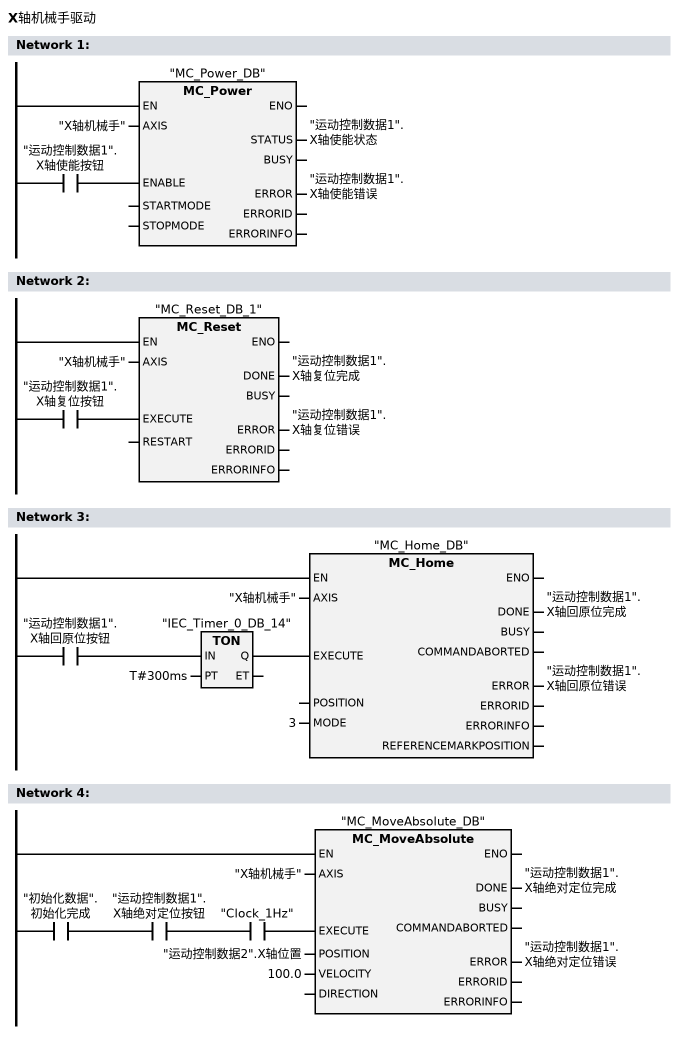
   "MC_Power_DB"(Axis := "X轴机械手",   // MC_Power
                 Enable := "运动控制数据1".X轴使能按钮,
                 Status => "运动控制数据1".X轴使能状态,
                 Error => "运动控制数据1".X轴使能错误);
END_REGION

REGION Network 2
   "MC_Reset_DB_1"(Axis := "X轴机械手",   // MC_Reset
                   Execute := "运动控制数据1".X轴复位按钮,
                   Done => "运动控制数据1".X轴复位完成,
                   Error => "运动控制数据1".X轴复位错误);
END_REGION

REGION Network 3
   "IEC_Timer_0_DB_14".TON(IN := "运动控制数据1".X轴回原位按钮, PT := T#300ms);
   "MC_Home_DB"(Axis := "X轴机械手",   // MC_Home
                Execute := "IEC_Timer_0_DB_14".Q,
                Mode := 3,
                Done => "运动控制数据1".X轴回原位完成,
                Error => "运动控制数据1".X轴回原位错误);
END_REGION

REGION Network 4
   "MC_MoveAbsolute_DB"(Axis := "X轴机械手",   // MC_MoveAbsolute
                        Execute := "初始化数据".初始化完成 AND "运动控制数据1".X轴绝对定位按钮 AND "Clock_1Hz",
                        Position := "运动控制数据2".X轴位置,
                        Velocity := 100.0,
                        Done => "运动控制数据1".X轴绝对定位完成,
                        Error => "运动控制数据1".X轴绝对定位错误);
END_REGION
END_FUNCTION

FUNCTION "Y轴机械手驱动" : Void   // FC2, LAD
{ S7_Optimized_Access := 'TRUE' }
VERSION : 0.1
BEGIN

REGION Network 1
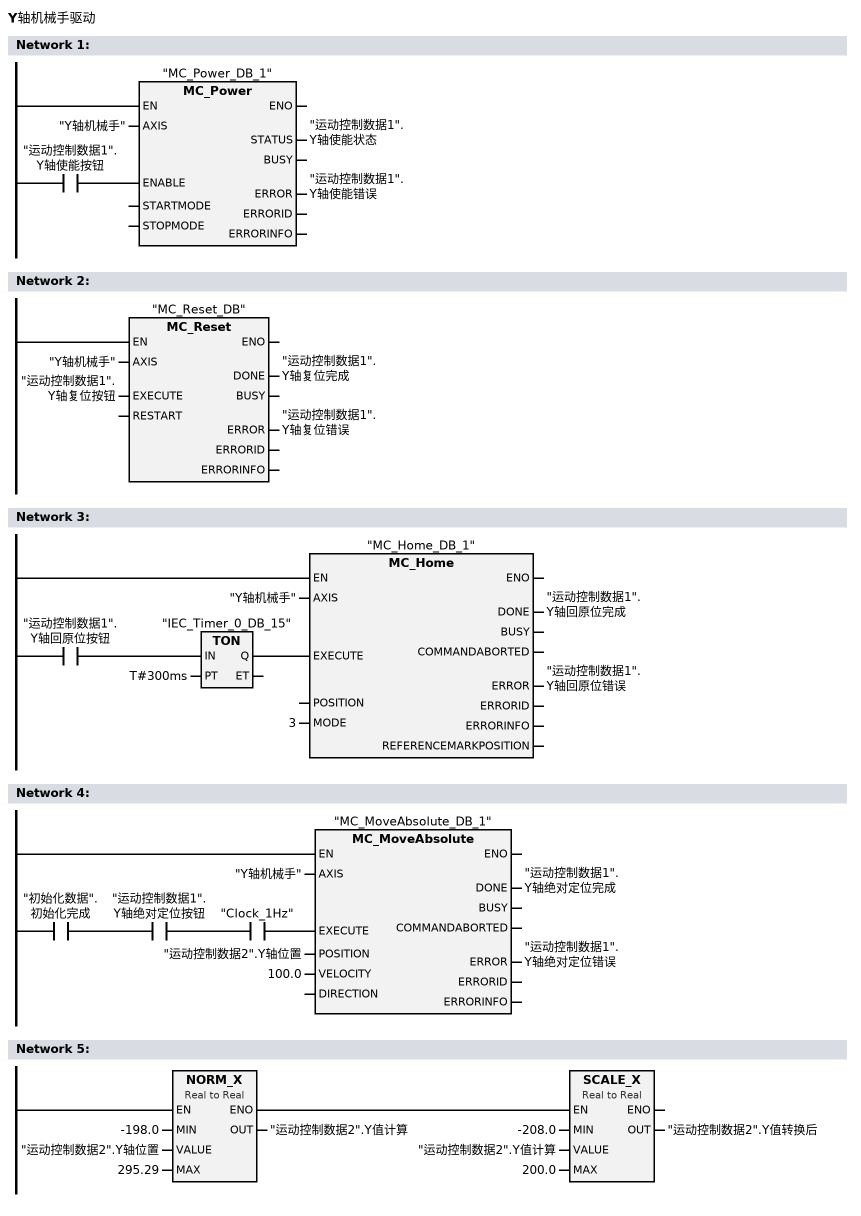
   "MC_Power_DB_1"(Axis := "Y轴机械手",   // MC_Power
                   Enable := "运动控制数据1".Y轴使能按钮,
                   Status => "运动控制数据1".Y轴使能状态,
                   Error => "运动控制数据1".Y轴使能错误);
END_REGION

REGION Network 2
   "MC_Reset_DB"(Axis := "Y轴机械手",   // MC_Reset
                 Execute := "运动控制数据1".Y轴复位按钮,
                 Done => "运动控制数据1".Y轴复位完成,
                 Error => "运动控制数据1".Y轴复位错误);
END_REGION

REGION Network 3
   "IEC_Timer_0_DB_15".TON(IN := "运动控制数据1".Y轴回原位按钮, PT := T#300ms);
   "MC_Home_DB_1"(Axis := "Y轴机械手",   // MC_Home
                  Execute := "IEC_Timer_0_DB_15".Q,
                  Mode := 3,
                  Done => "运动控制数据1".Y轴回原位完成,
                  Error => "运动控制数据1".Y轴回原位错误);
END_REGION

REGION Network 4
   "MC_MoveAbsolute_DB_1"(Axis := "Y轴机械手",   // MC_MoveAbsolute
                          Execute := "初始化数据".初始化完成 AND "运动控制数据1".Y轴绝对定位按钮 AND "Clock_1Hz",
                          Position := "运动控制数据2".Y轴位置,
                          Velocity := 100.0,
                          Done => "运动控制数据1".Y轴绝对定位完成,
                          Error => "运动控制数据1".Y轴绝对定位错误);
END_REGION

REGION Network 5
   RUNG wire#powerrail
      { S7_Templates := "[SrcType := Real, DestType := Real]" } Normalize(min := -198.0, value := "运动控制数据2".Y轴位置, max := 295.29, out => "运动控制数据2".Y值计算)
      { S7_Templates := "[SrcType := Real, DestType := Real]" } Scale(min := -208.0, value := "运动控制数据2".Y值计算, max := 200.0, out => "运动控制数据2".Y值转换后)
   END_RUNG
   // the same network as SCL:
   "运动控制数据2".Y值计算 := NORM_X(MIN := -198.0, VALUE := "运动控制数据2".Y轴位置, MAX := 295.29);
   "运动控制数据2".Y值转换后 := SCALE_X(MIN := -208.0, VALUE := "运动控制数据2".Y值计算, MAX := 200.0);
END_REGION
END_FUNCTION

FUNCTION "传输皮带" : Void   // FC3, LAD
{ S7_Optimized_Access := 'TRUE' }
VERSION : 0.1
BEGIN

REGION Network 1
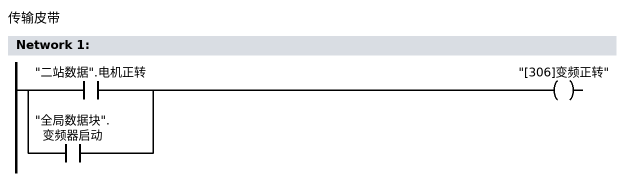
   RUNG wire#powerrail
      Contact( "二站数据".电机正转 )
      wire#w1
      Coil( "[306]变频正转" )
   END_RUNG
   RUNG wire#powerrail
      Contact( "全局数据块".变频器启动 )
   END_RUNG wire#w1
   // the same network as SCL:
   "[306]变频正转" := "二站数据".电机正转 OR "全局数据块".变频器启动;
END_REGION
END_FUNCTION

FUNCTION "00.轴初始化程序" : Void   // FC11, LAD
{ S7_Optimized_Access := 'TRUE' }
VERSION : 0.1
   VAR_TEMP   // added for the SCL form of the ladder/FBD networks
      _w1 : Bool;
   END_VAR
BEGIN

REGION Network 1
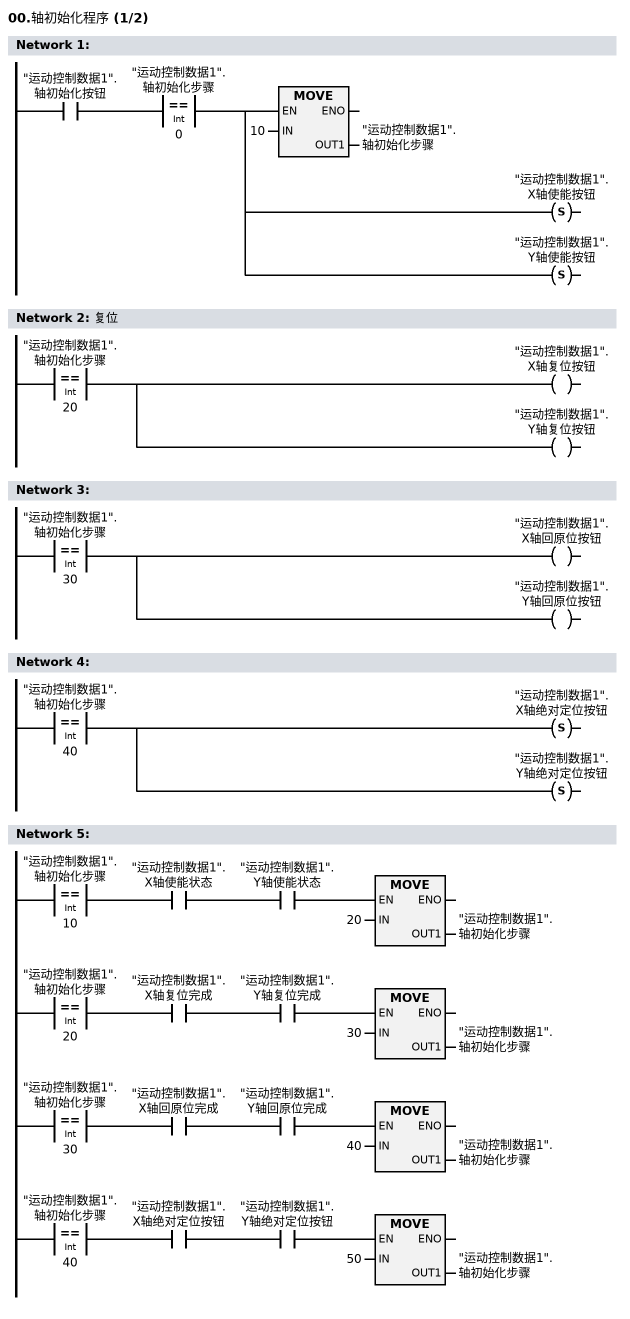
   RUNG wire#powerrail
      Contact( "运动控制数据1".轴初始化按钮 )
      { S7_Templates := "SrcType := Int" } EQ_Contact(in1 := "运动控制数据1".轴初始化步骤, in2 := 0)
      wire#w1
      Move(in := 10, out1 => "运动控制数据1".轴初始化步骤)
   END_RUNG
   RUNG wire#w1
      S_Coil( "运动控制数据1".X轴使能按钮 )
   END_RUNG
   RUNG wire#w1
      S_Coil( "运动控制数据1".Y轴使能按钮 )
   END_RUNG
   // the same network as SCL:
   #_w1 := "运动控制数据1".轴初始化按钮 AND ("运动控制数据1".轴初始化步骤 = 0);
   IF #_w1 THEN
       "运动控制数据1".轴初始化步骤 := 10;
       "运动控制数据1".X轴使能按钮 := TRUE;
       "运动控制数据1".Y轴使能按钮 := TRUE;
   END_IF;
END_REGION

REGION Network 2: 复位
   RUNG wire#powerrail
      { S7_Templates := "SrcType := Int" } EQ_Contact(in1 := "运动控制数据1".轴初始化步骤, in2 := 20)
      wire#w1
      Coil( "运动控制数据1".X轴复位按钮 )
   END_RUNG
   RUNG wire#w1
      Coil( "运动控制数据1".Y轴复位按钮 )
   END_RUNG
   // the same network as SCL:
   "运动控制数据1".X轴复位按钮 := "运动控制数据1".轴初始化步骤 = 20;
   "运动控制数据1".Y轴复位按钮 := "运动控制数据1".X轴复位按钮;
END_REGION

REGION Network 3
   RUNG wire#powerrail
      { S7_Templates := "SrcType := Int" } EQ_Contact(in1 := "运动控制数据1".轴初始化步骤, in2 := 30)
      wire#w1
      Coil( "运动控制数据1".X轴回原位按钮 )
   END_RUNG
   RUNG wire#w1
      Coil( "运动控制数据1".Y轴回原位按钮 )
   END_RUNG
   // the same network as SCL:
   "运动控制数据1".X轴回原位按钮 := "运动控制数据1".轴初始化步骤 = 30;
   "运动控制数据1".Y轴回原位按钮 := "运动控制数据1".X轴回原位按钮;
END_REGION

REGION Network 4
   RUNG wire#powerrail
      { S7_Templates := "SrcType := Int" } EQ_Contact(in1 := "运动控制数据1".轴初始化步骤, in2 := 40)
      wire#w1
      S_Coil( "运动控制数据1".X轴绝对定位按钮 )
   END_RUNG
   RUNG wire#w1
      S_Coil( "运动控制数据1".Y轴绝对定位按钮 )
   END_RUNG
   // the same network as SCL:
   IF "运动控制数据1".轴初始化步骤 = 40 THEN
       "运动控制数据1".X轴绝对定位按钮 := TRUE;
       "运动控制数据1".Y轴绝对定位按钮 := TRUE;
   END_IF;
END_REGION

REGION Network 5
   RUNG wire#powerrail
      { S7_Templates := "SrcType := Int" } EQ_Contact(in1 := "运动控制数据1".轴初始化步骤, in2 := 10)
      Contact( "运动控制数据1".X轴使能状态 )
      Contact( "运动控制数据1".Y轴使能状态 )
      Move(in := 20, out1 => "运动控制数据1".轴初始化步骤)
   END_RUNG
   RUNG wire#powerrail
      { S7_Templates := "SrcType := Int" } EQ_Contact(in1 := "运动控制数据1".轴初始化步骤, in2 := 20)
      Contact( "运动控制数据1".X轴复位完成 )
      Contact( "运动控制数据1".Y轴复位完成 )
      Move(in := 30, out1 => "运动控制数据1".轴初始化步骤)
   END_RUNG
   RUNG wire#powerrail
      { S7_Templates := "SrcType := Int" } EQ_Contact(in1 := "运动控制数据1".轴初始化步骤, in2 := 30)
      Contact( "运动控制数据1".X轴回原位完成 )
      Contact( "运动控制数据1".Y轴回原位完成 )
      Move(in := 40, out1 => "运动控制数据1".轴初始化步骤)
   END_RUNG
   RUNG wire#powerrail
      { S7_Templates := "SrcType := Int" } EQ_Contact(in1 := "运动控制数据1".轴初始化步骤, in2 := 40)
      Contact( "运动控制数据1".X轴绝对定位按钮 )
      Contact( "运动控制数据1".Y轴绝对定位按钮 )
      Move(in := 50, out1 => "运动控制数据1".轴初始化步骤)
   END_RUNG
   // the same network as SCL:
   IF ("运动控制数据1".轴初始化步骤 = 10) AND "运动控制数据1".X轴使能状态 AND "运动控制数据1".Y轴使能状态 THEN "运动控制数据1".轴初始化步骤 := 20; END_IF;
   IF ("运动控制数据1".轴初始化步骤 = 20) AND "运动控制数据1".X轴复位完成 AND "运动控制数据1".Y轴复位完成 THEN "运动控制数据1".轴初始化步骤 := 30; END_IF;
   IF ("运动控制数据1".轴初始化步骤 = 30) AND "运动控制数据1".X轴回原位完成 AND "运动控制数据1".Y轴回原位完成 THEN
       "运动控制数据1".轴初始化步骤 := 40;
   END_IF;
   IF ("运动控制数据1".轴初始化步骤 = 40) AND "运动控制数据1".X轴绝对定位按钮 AND "运动控制数据1".Y轴绝对定位按钮 THEN
       "运动控制数据1".轴初始化步骤 := 50;
   END_IF;
END_REGION

REGION Network 6: 轴初始化完成
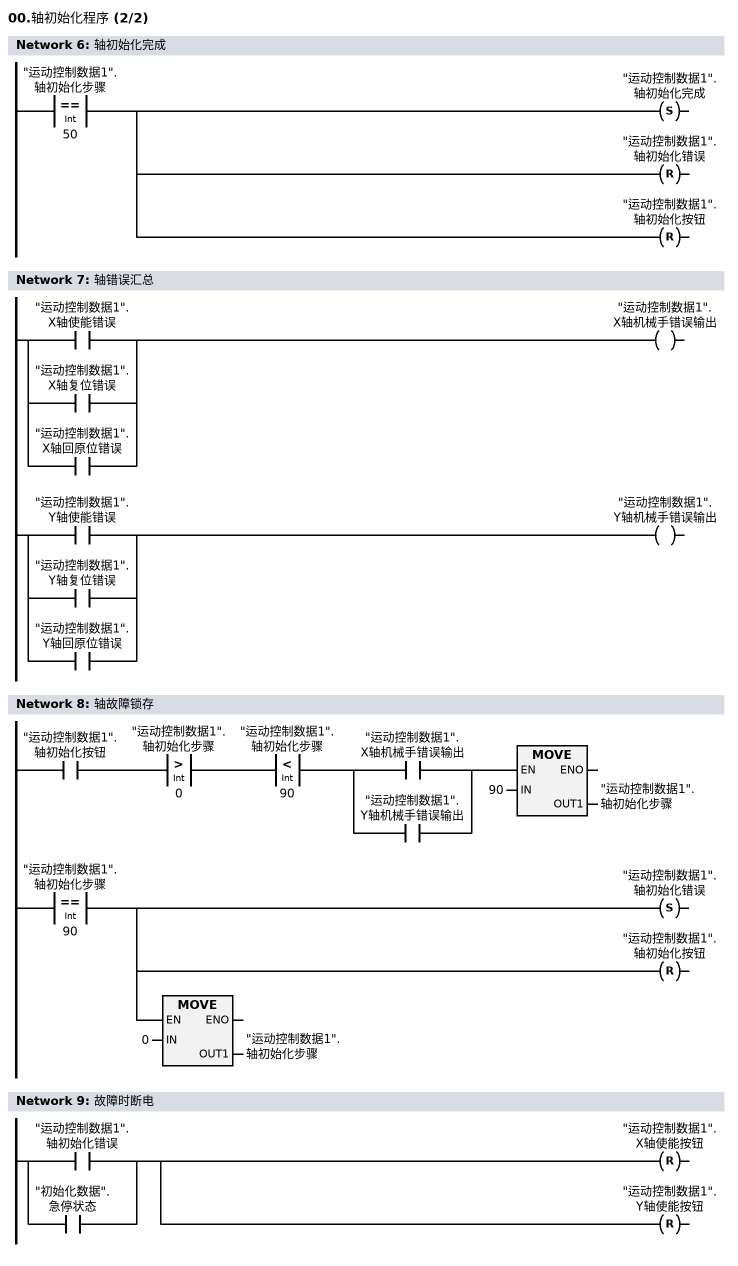
   RUNG wire#powerrail
      { S7_Templates := "SrcType := Int" } EQ_Contact(in1 := "运动控制数据1".轴初始化步骤, in2 := 50)
      wire#w1
      S_Coil( "运动控制数据1".轴初始化完成 )
   END_RUNG
   RUNG wire#w1
      R_Coil( "运动控制数据1".轴初始化错误 )
   END_RUNG
   RUNG wire#w1
      R_Coil( "运动控制数据1".轴初始化按钮 )
   END_RUNG
   // the same network as SCL:
   IF "运动控制数据1".轴初始化步骤 = 50 THEN
       "运动控制数据1".轴初始化完成 := TRUE;
       "运动控制数据1".轴初始化错误 := FALSE;
       "运动控制数据1".轴初始化按钮 := FALSE;
   END_IF;
END_REGION

REGION Network 7: 轴错误汇总
   RUNG wire#powerrail
      Contact( "运动控制数据1".X轴使能错误 )
      wire#w1
      Coil( "运动控制数据1".X轴机械手错误输出 )
   END_RUNG
   RUNG wire#powerrail
      Contact( "运动控制数据1".X轴复位错误 )
   END_RUNG wire#w1
   RUNG wire#powerrail
      Contact( "运动控制数据1".X轴回原位错误 )
   END_RUNG wire#w1
   RUNG wire#powerrail
      Contact( "运动控制数据1".Y轴使能错误 )
      wire#w2
      Coil( "运动控制数据1".Y轴机械手错误输出 )
   END_RUNG
   RUNG wire#powerrail
      Contact( "运动控制数据1".Y轴复位错误 )
   END_RUNG wire#w2
   RUNG wire#powerrail
      Contact( "运动控制数据1".Y轴回原位错误 )
   END_RUNG wire#w2
   // the same network as SCL:
   "运动控制数据1".X轴机械手错误输出 := "运动控制数据1".X轴使能错误 OR "运动控制数据1".X轴复位错误 OR "运动控制数据1".X轴回原位错误;
   "运动控制数据1".Y轴机械手错误输出 := "运动控制数据1".Y轴使能错误 OR "运动控制数据1".Y轴复位错误 OR "运动控制数据1".Y轴回原位错误;
END_REGION

REGION Network 8: 轴故障锁存
   RUNG wire#powerrail
      Contact( "运动控制数据1".轴初始化按钮 )
      { S7_Templates := "SrcType := Int" } GT_Contact(in1 := "运动控制数据1".轴初始化步骤, in2 := 0)
      { S7_Templates := "SrcType := Int" } LT_Contact(in1 := "运动控制数据1".轴初始化步骤, in2 := 90)
      wire#w1
      Contact( "运动控制数据1".X轴机械手错误输出 )
      wire#w2
      Move(in := 90, out1 => "运动控制数据1".轴初始化步骤)
   END_RUNG
   RUNG wire#w1
      Contact( "运动控制数据1".Y轴机械手错误输出 )
   END_RUNG wire#w2
   RUNG wire#powerrail
      { S7_Templates := "SrcType := Int" } EQ_Contact(in1 := "运动控制数据1".轴初始化步骤, in2 := 90)
      wire#w3
      S_Coil( "运动控制数据1".轴初始化错误 )
   END_RUNG
   RUNG wire#w3
      R_Coil( "运动控制数据1".轴初始化按钮 )
   END_RUNG
   RUNG wire#w3
      Move(in := 0, out1 => "运动控制数据1".轴初始化步骤)
   END_RUNG
   // the same network as SCL:
   IF "运动控制数据1".轴初始化按钮 AND ("运动控制数据1".轴初始化步骤 > 0) AND ("运动控制数据1".轴初始化步骤 < 90) AND ("运动控制数据1".X轴机械手错误输出 OR "运动控制数据1".Y轴机械手错误输出) THEN
       "运动控制数据1".轴初始化步骤 := 90;
   END_IF;
   IF "运动控制数据1".轴初始化步骤 = 90 THEN
       "运动控制数据1".轴初始化错误 := TRUE;
       "运动控制数据1".轴初始化按钮 := FALSE;
       "运动控制数据1".轴初始化步骤 := 0;
   END_IF;
END_REGION

REGION Network 9: 故障时断电
   RUNG wire#powerrail
      Contact( "运动控制数据1".轴初始化错误 )
      wire#w1
      R_Coil( "运动控制数据1".X轴使能按钮 )
   END_RUNG
   RUNG wire#powerrail
      Contact( "初始化数据".急停状态 )
   END_RUNG wire#w1
   RUNG wire#w1
      R_Coil( "运动控制数据1".Y轴使能按钮 )
   END_RUNG
   // the same network as SCL:
   IF "运动控制数据1".轴初始化错误 OR "初始化数据".急停状态 THEN
       "运动控制数据1".X轴使能按钮 := FALSE;
       "运动控制数据1".Y轴使能按钮 := FALSE;
   END_IF;
END_REGION
END_FUNCTION

// folder: 通讯模块

FUNCTION "产线通讯" : Void   // FC4, LAD
{ S7_Optimized_Access := 'TRUE' }
VERSION : 0.1
BEGIN

REGION Network 1: 心跳
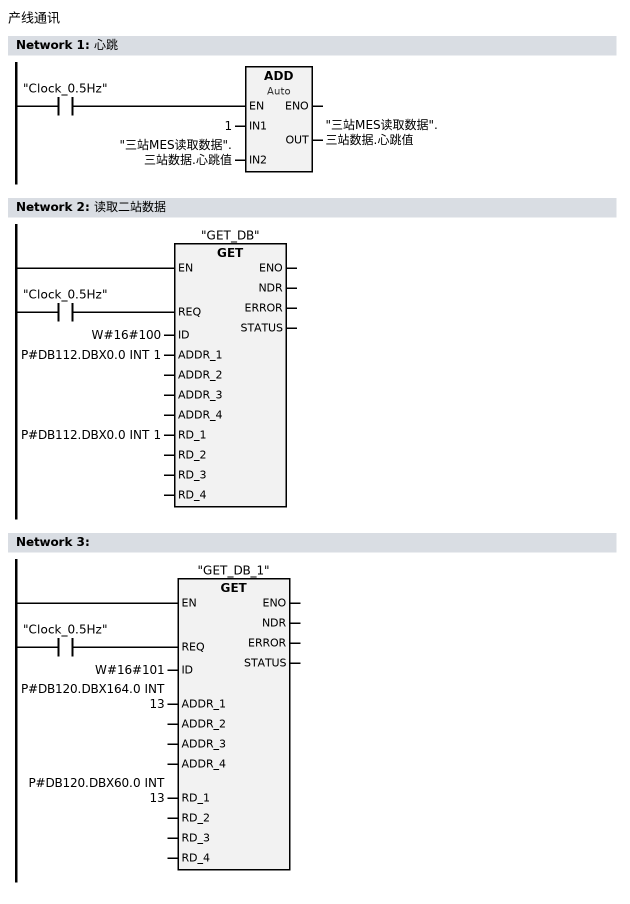
   RUNG wire#powerrail
      Contact( "Clock_0.5Hz" )
      Add(in1 := 1, in2 := "三站MES读取数据".三站数据.心跳值, out => "三站MES读取数据".三站数据.心跳值)
   END_RUNG
   // the same network as SCL:
   IF "Clock_0.5Hz" THEN "三站MES读取数据".三站数据.心跳值 := 1 + "三站MES读取数据".三站数据.心跳值; END_IF;
END_REGION

REGION Network 2: 读取二站数据
   "GET_DB"(REQ := "Clock_0.5Hz", ID := W#16#100, ADDR_1 := P#DB112.DBX0.0 INT 1, RD_1 := P#DB112.DBX0.0 INT 1);   // GET
END_REGION

REGION Network 3
   "GET_DB_1"(REQ := "Clock_0.5Hz",   // GET
              ID := W#16#101,
              ADDR_1 := P#DB120.DBX164.0 INT 13,
              RD_1 := P#DB120.DBX60.0 INT 13);
END_REGION
END_FUNCTION

FUNCTION "称重器通讯" : Void   // FC10, LAD
{ S7_Optimized_Access := 'TRUE' }
VERSION : 0.1
BEGIN

REGION Network 1
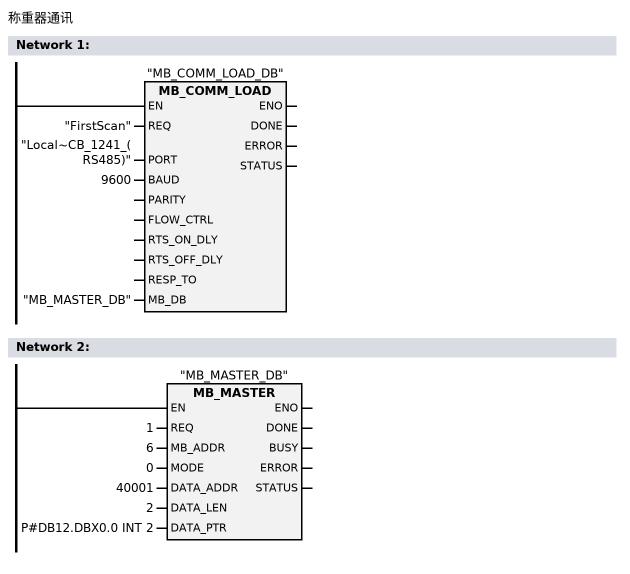
   "MB_COMM_LOAD_DB"(REQ := "FirstScan", PORT := "Local~CB_1241_(RS485)", BAUD := 9600, MB_DB := "MB_MASTER_DB");   // MB_COMM_LOAD
END_REGION

REGION Network 2
   "MB_MASTER_DB"(REQ := 1,   // MB_MASTER
                  MB_ADDR := 6,
                  MODE := 0,
                  DATA_ADDR := 40001,
                  DATA_LEN := 2,
                  DATA_PTR := P#DB12.DBX0.0 INT 2);
END_REGION
END_FUNCTION

FUNCTION "AI视觉信号映射" : Void   // FC12, LAD
{ S7_Optimized_Access := 'TRUE' }
VERSION : 0.1
BEGIN

REGION Network 1
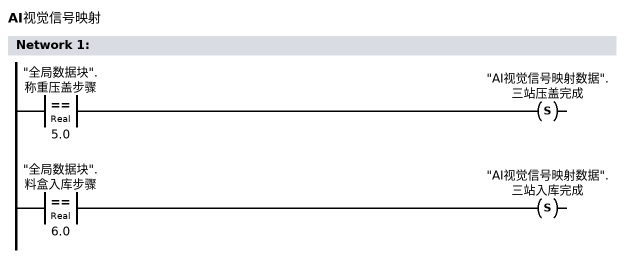
   RUNG wire#powerrail
      { S7_Templates := "SrcType := Real" } EQ_Contact(in1 := "全局数据块".称重压盖步骤, in2 := 5.0)
      S_Coil( "AI视觉信号映射数据".三站压盖完成 )
   END_RUNG
   RUNG wire#powerrail
      { S7_Templates := "SrcType := Real" } EQ_Contact(in1 := "全局数据块".料盒入库步骤, in2 := 6.0)
      S_Coil( "AI视觉信号映射数据".三站入库完成 )
   END_RUNG
   // the same network as SCL:
   IF "全局数据块".称重压盖步骤 = 5.0 THEN "AI视觉信号映射数据".三站压盖完成 := TRUE; END_IF;
   IF "全局数据块".料盒入库步骤 = 6.0 THEN "AI视觉信号映射数据".三站入库完成 := TRUE; END_IF;
END_REGION
END_FUNCTION

FUNCTION "扫码器通讯" : Void   // FC13, LAD
{ S7_Optimized_Access := 'TRUE' }
VERSION : 0.1
BEGIN

REGION Network 1: 入站扫码器
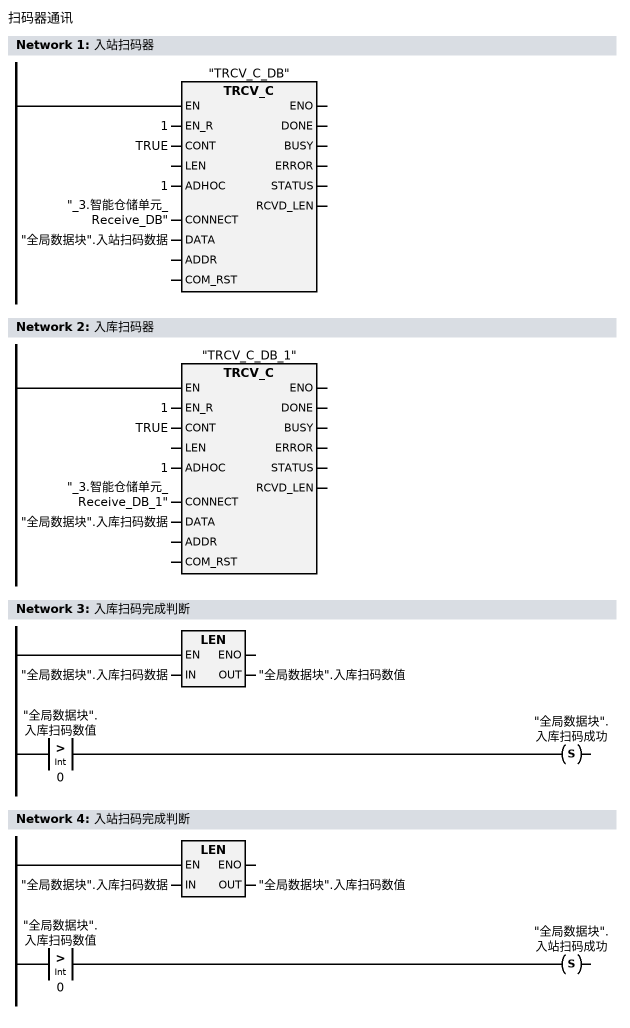
   "TRCV_C_DB"(EN_R := 1, CONT := TRUE, ADHOC := 1, CONNECT := "_3.智能仓储单元_Receive_DB", DATA := "全局数据块".入站扫码数据);   // TRCV_C
END_REGION

REGION Network 2: 入库扫码器
   "TRCV_C_DB_1"(EN_R := 1,   // TRCV_C
                 CONT := TRUE,
                 ADHOC := 1,
                 CONNECT := "_3.智能仓储单元_Receive_DB_1",
                 DATA := "全局数据块".入库扫码数据);
END_REGION

REGION Network 3: 入库扫码完成判断
   "全局数据块".入库扫码数值 := LEN(IN := "全局数据块".入库扫码数据);
   IF "全局数据块".入库扫码数值 > 0 THEN "全局数据块".入库扫码成功 := TRUE; END_IF;
END_REGION

REGION Network 4: 入站扫码完成判断
   "全局数据块".入库扫码数值 := LEN(IN := "全局数据块".入库扫码数据);
   IF "全局数据块".入库扫码数值 > 0 THEN "全局数据块".入站扫码成功 := TRUE; END_IF;
END_REGION
END_FUNCTION

FUNCTION "虚拟联动映射" : Void   // FC15, LAD
{ S7_Optimized_Access := 'TRUE' }
VERSION : 0.1
BEGIN

REGION Network 1
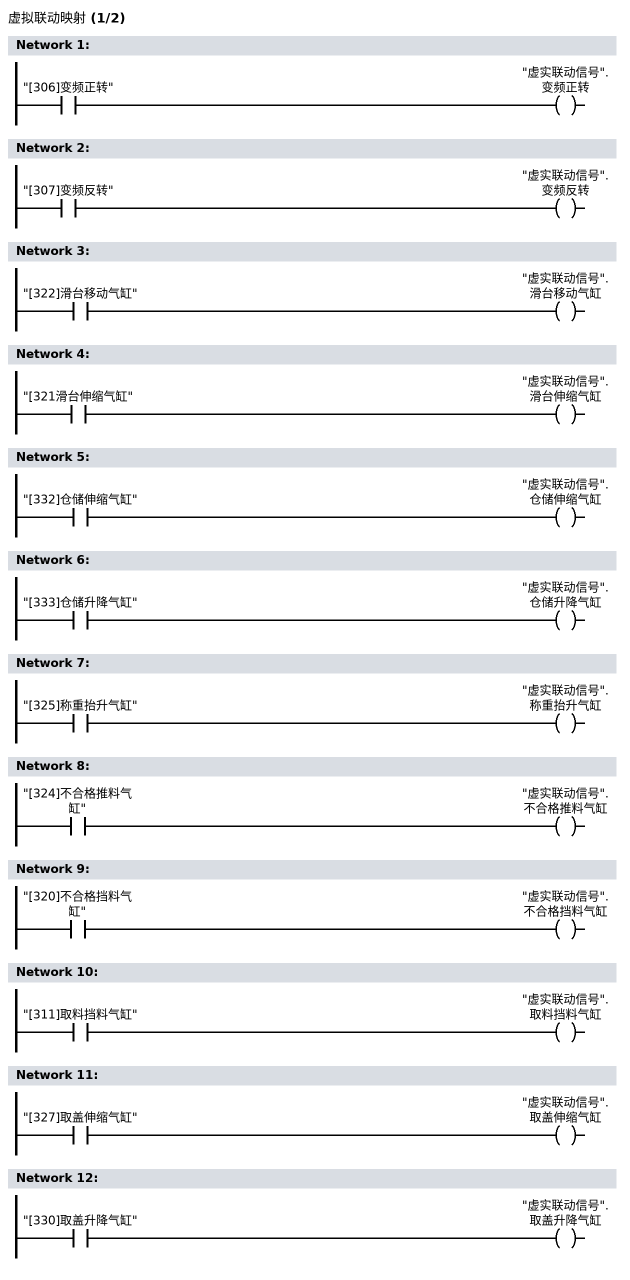
   RUNG wire#powerrail
      Contact( "[306]变频正转" )
      Coil( "虚实联动信号".变频正转 )
   END_RUNG
   // the same network as SCL:
   "虚实联动信号".变频正转 := "[306]变频正转";
END_REGION

REGION Network 2
   RUNG wire#powerrail
      Contact( "[307]变频反转" )
      Coil( "虚实联动信号".变频反转 )
   END_RUNG
   // the same network as SCL:
   "虚实联动信号".变频反转 := "[307]变频反转";
END_REGION

REGION Network 3
   RUNG wire#powerrail
      Contact( "[322]滑台移动气缸" )
      Coil( "虚实联动信号".滑台移动气缸 )
   END_RUNG
   // the same network as SCL:
   "虚实联动信号".滑台移动气缸 := "[322]滑台移动气缸";
END_REGION

REGION Network 4
   RUNG wire#powerrail
      Contact( "[321滑台伸缩气缸" )
      Coil( "虚实联动信号".滑台伸缩气缸 )
   END_RUNG
   // the same network as SCL:
   "虚实联动信号".滑台伸缩气缸 := "[321滑台伸缩气缸";
END_REGION

REGION Network 5
   RUNG wire#powerrail
      Contact( "[332]仓储伸缩气缸" )
      Coil( "虚实联动信号".仓储伸缩气缸 )
   END_RUNG
   // the same network as SCL:
   "虚实联动信号".仓储伸缩气缸 := "[332]仓储伸缩气缸";
END_REGION

REGION Network 6
   RUNG wire#powerrail
      Contact( "[333]仓储升降气缸" )
      Coil( "虚实联动信号".仓储升降气缸 )
   END_RUNG
   // the same network as SCL:
   "虚实联动信号".仓储升降气缸 := "[333]仓储升降气缸";
END_REGION

REGION Network 7
   RUNG wire#powerrail
      Contact( "[325]称重抬升气缸" )
      Coil( "虚实联动信号".称重抬升气缸 )
   END_RUNG
   // the same network as SCL:
   "虚实联动信号".称重抬升气缸 := "[325]称重抬升气缸";
END_REGION

REGION Network 8
   RUNG wire#powerrail
      Contact( "[324]不合格推料气缸" )
      Coil( "虚实联动信号".不合格推料气缸 )
   END_RUNG
   // the same network as SCL:
   "虚实联动信号".不合格推料气缸 := "[324]不合格推料气缸";
END_REGION

REGION Network 9
   RUNG wire#powerrail
      Contact( "[320]不合格挡料气缸" )
      Coil( "虚实联动信号".不合格挡料气缸 )
   END_RUNG
   // the same network as SCL:
   "虚实联动信号".不合格挡料气缸 := "[320]不合格挡料气缸";
END_REGION

REGION Network 10
   RUNG wire#powerrail
      Contact( "[311]取料挡料气缸" )
      Coil( "虚实联动信号".取料挡料气缸 )
   END_RUNG
   // the same network as SCL:
   "虚实联动信号".取料挡料气缸 := "[311]取料挡料气缸";
END_REGION

REGION Network 11
   RUNG wire#powerrail
      Contact( "[327]取盖伸缩气缸" )
      Coil( "虚实联动信号".取盖伸缩气缸 )
   END_RUNG
   // the same network as SCL:
   "虚实联动信号".取盖伸缩气缸 := "[327]取盖伸缩气缸";
END_REGION

REGION Network 12
   RUNG wire#powerrail
      Contact( "[330]取盖升降气缸" )
      Coil( "虚实联动信号".取盖升降气缸 )
   END_RUNG
   // the same network as SCL:
   "虚实联动信号".取盖升降气缸 := "[330]取盖升降气缸";
END_REGION

REGION Network 13
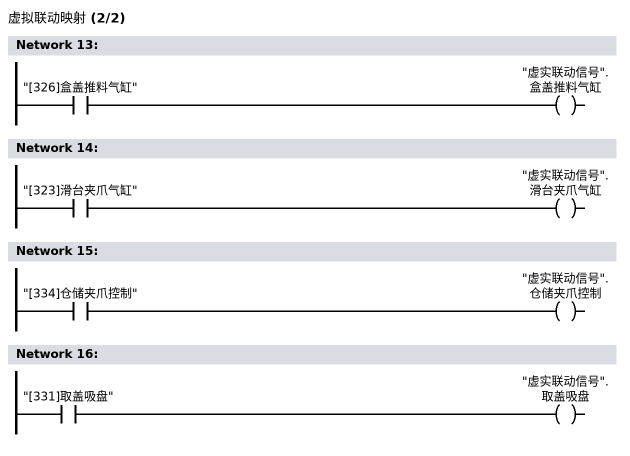
   RUNG wire#powerrail
      Contact( "[326]盒盖推料气缸" )
      Coil( "虚实联动信号".盒盖推料气缸 )
   END_RUNG
   // the same network as SCL:
   "虚实联动信号".盒盖推料气缸 := "[326]盒盖推料气缸";
END_REGION

REGION Network 14
   RUNG wire#powerrail
      Contact( "[323]滑台夹爪气缸" )
      Coil( "虚实联动信号".滑台夹爪气缸 )
   END_RUNG
   // the same network as SCL:
   "虚实联动信号".滑台夹爪气缸 := "[323]滑台夹爪气缸";
END_REGION

REGION Network 15
   RUNG wire#powerrail
      Contact( "[334]仓储夹爪控制" )
      Coil( "虚实联动信号".仓储夹爪控制 )
   END_RUNG
   // the same network as SCL:
   "虚实联动信号".仓储夹爪控制 := "[334]仓储夹爪控制";
END_REGION

REGION Network 16
   RUNG wire#powerrail
      Contact( "[331]取盖吸盘" )
      Coil( "虚实联动信号".取盖吸盘 )
   END_RUNG
   // the same network as SCL:
   "虚实联动信号".取盖吸盘 := "[331]取盖吸盘";
END_REGION
END_FUNCTION

FUNCTION "数据转换检测" : Void   // FC17, LAD
{ S7_Optimized_Access := 'TRUE' }
VERSION : 0.1
BEGIN
END_FUNCTION

FUNCTION "MES数据映射" : Void   // FC18, LAD
{ S7_Optimized_Access := 'TRUE' }
VERSION : 0.1
BEGIN
END_FUNCTION

// ===== PLC "0.数据管理单元"  CPU 1511-1 PN =====

VAR_GLOBAL   // PLC tag table "默认变量表"
   "System_Byte" AT %MB501 : Byte;
   "FirstScan" AT %M501.0 : Bool;
   "DiagStatusUpdate" AT %M501.1 : Bool;
   "AlwaysTRUE" AT %M501.2 : Bool;
   "AlwaysFALSE" AT %M501.3 : Bool;
   "Clock_Byte" AT %MB500 : Byte;
   "Clock_10Hz" AT %M500.0 : Bool;
   "Clock_5Hz" AT %M500.1 : Bool;
   "Clock_2.5Hz" AT %M500.2 : Bool;
   "Clock_2Hz" AT %M500.3 : Bool;
   "Clock_1.25Hz" AT %M500.4 : Bool;
   "Clock_1Hz" AT %M500.5 : Bool;
   "Clock_0.625Hz" AT %M500.6 : Bool;
   "Clock_0.5Hz" AT %M500.7 : Bool;
   "Tag_1" AT %M12.0 : Bool;
END_VAR

VAR_GLOBAL   // PLC tag table "数据管理单元变量表"
   "[100]启动按钮" AT %I0.0 : Bool;
   "[101]停止按钮" AT %I0.1 : Bool;
   "[102]复位按钮" AT %I0.2 : Bool;
   "[103]急停按钮" AT %I0.3 : Bool;
   "[104]手/自动" AT %I0.4 : Bool;
   "读取电压" AT %ID134 : DWord;
   "读取电流" AT %ID138 : DWord;
   "读取有功功率" AT %ID142 : DWord;
   "读取无功功率" AT %ID146 : DWord;
   "读取视在功率" AT %ID150 : DWord;
   "读取功率因数" AT %ID154 : DWord;
   "读取保留参数" AT %ID158 : DWord;
   "读取电网频率" AT %ID162 : DWord;
   "读取总电能" AT %ID170 : DWord;
   "读取温度" AT %IW190 : Int;
   "读取湿度" AT %IW192 : Int;
   "[105]允许下单" AT %I0.7 : Bool;
   "[156]安全光栅" AT %I5.6 : Bool;
   "[300]黄色灯" AT %Q0.0 : Bool;
   "[301]绿色灯" AT %Q0.1 : Bool;
   "[302]红色灯" AT %Q0.2 : Bool;
   "写入电能清零" AT %QW180 : Word;
   "[320]LORA-黄灯" AT %Q2.0 : Bool;
   "[340]LORA-绿灯" AT %Q4.0 : Bool;
   "[360]LORA-红灯" AT %Q6.0 : Bool;
   "Tag_2" AT %Q2.1 : Bool;
   "[303]绿色指示灯" AT %Q0.3 : Bool;
   "[304]红色指示灯" AT %Q0.4 : Bool;
   "[307]声光报警" AT %Q0.7 : Bool;
END_VAR

DATA_BLOCK "订单信息下发_DB"   // DB4
{ S7_Optimized_Access := 'TRUE' }
VERSION : 0.1
// stored: InstanceOfName 订单信息下发
"订单信息下发"
BEGIN
END_DATA_BLOCK

DATA_BLOCK "MES订单数据"   // DB121
{ S7_Optimized_Access := 'FALSE' }
VERSION : 0.1
   VAR
      订单ID : Int;
      AB物料 : Int;
      "8mm钢珠数量" : Int;
      "10mm钢珠数量" : Int;
      存储仓位 : Int;
      PLC通讯心跳 : Int;
      MES下单请求 : Bool;
      PLC订单已下发 : Bool;
      产线可接单 : Bool;
      订单已完成 : Bool;
      完成订单ID : Int;
   END_VAR
BEGIN
END_DATA_BLOCK

// folder: System blocks/Program resources

DATA_BLOCK "IEC_Timer_0_DB"   // DB2
{ S7_Optimized_Access := 'TRUE' }
AUTHOR : Simatic
FAMILY : IEC
NAME : IEC_TMR
VERSION : 1.0
// stored: InstanceOfName IEC_TIMER
"IEC_TIMER"
BEGIN
END_DATA_BLOCK

DATA_BLOCK "IEC_Timer_0_DB_1"   // DB5
{ S7_Optimized_Access := 'TRUE' }
AUTHOR : Simatic
FAMILY : IEC
NAME : IEC_TMR
VERSION : 1.0
// stored: InstanceOfName IEC_TIMER
"IEC_TIMER"
BEGIN
END_DATA_BLOCK

// folder: 通讯数据

DATA_BLOCK "初始化数据"   // DB1
{ S7_Optimized_Access := 'FALSE' }
VERSION : 0.1
   VAR
      手动模式 : Bool;
      自动模式 : Bool;
      自动运行模式 : Bool;
      产线复位步骤 : Int;
      急停状态 : Bool;
      红灯_内部 : Bool;
      黄灯_内部 : Bool;
      绿灯_内部 : Bool;
      报警等级 : Int;
      报警确认按钮 : Bool;
      初始化完成 : Bool;
   END_VAR
BEGIN
END_DATA_BLOCK

DATA_BLOCK "全局数据"   // DB3
{ S7_Optimized_Access := 'FALSE' }
VERSION : 0.1
   VAR
      产线状态正常 : Bool;
      产线三站空闲 : Bool;
      产线复位按钮 : Bool;
      触摸屏下单按钮 : Bool;
      触摸屏复位按钮 : Bool;
      复位上升沿 : Bool;
      产线正在运行 : Bool;
   END_VAR
BEGIN
END_DATA_BLOCK

DATA_BLOCK "0.MES通讯数据"   // DB120
{ S7_Optimized_Access := 'FALSE' }
VERSION : 0.1
   VAR
      一站数据 : Struct
         在线状态 : Int;
         运行模式 : Int;   // 0 手动 / 1 自动待机 / 2 自动运行
         忙碌状态 : Int;   // 0 空闲 / 1 忙碌
         故障状态 : Int;   // 0 = 无故障
         当前订单ID : Int;   // 当前处理的订单
         当前步骤 : Real;
         心跳值 : Int;
         一站完成 : Bool;
         一站已接收 : Bool;
         保留_1 : Bool;
         保留_2 : Bool;
         保留_3 : Bool;
         保留_4 : Bool;
         保留_5 : Bool;
         保留_6 : Bool;
         扫码条码数据 : Int;
         转盘当前角度 : Real;
         机械手当前位置 : Real;
         深度检测值 : Real;
         料盒使用数 : Int;
         A料使用数 : Int;
         B料使用数 : Int;
         一站保留数据 : Array[0..9] of Int;
      END_STRUCT;
      二站数据 : Struct
         在线状态 : Int;
         运行模式 : Int;   // 0 手动 / 1 自动待机 / 2 自动运行
         忙碌状态 : Int;   // 0 空闲 / 1 忙碌
         故障状态 : Int;   // 0 = 无故障
         当前订单ID : Int;   // 当前处理的订单
         当前步骤 : Real;
         心跳值 : Int;
         二站完成 : Bool;
         二站已接收 : Bool;
         保留_1 : Bool;
         保留_2 : Bool;
         保留_3 : Bool;
         保留_4 : Bool;
         保留_5 : Bool;
         保留_6 : Bool;
         二站扫码数据 : Int;
         "8mm已灌注数量" : Int;
         "10mm已灌注数量" : Int;
         "8mml料仓钢珠有无" : Bool;   // 1有0无
         "10mm料仓钢珠有无" : Bool;   // 1有0无
         二站保留数据 : Array[0..9] of Int;
      END_STRUCT;
      三站数据 : Struct
         在线状态 : Int;
         运行模式 : Int;   // 0 手动 / 1 自动待机 / 2 自动运行
         忙碌状态 : Int;   // 0 空闲 / 1 忙碌
         故障状态 : Int;   // 0 = 无故障
         当前订单ID : Int;   // 当前处理的订单
         当前步骤 : Real;
         心跳值 : Int;
         三站完成 : Bool;
         三站已接收 : Bool;
         保留_1 : Bool;
         保留_2 : Bool;
         保留_3 : Bool;
         保留_4 : Bool;
         保留_5 : Bool;
         保留_6 : Bool;
         仓位状态 : Array[0..8] of Bool;
         入站扫码数据 : Int;
         入库扫码数据 : Int;
         称重数据 : Int;
         产品合格状态 : Int;
         合格产品计数 : Int;
         不合格产品计数 : Int;
         X轴当前位置 : Real;
         Y轴当前位置 : Real;
         完成订单ID : Int;
         三站保留数据 : Array[0..8] of Int;
      END_STRUCT;
      订单数据 : Struct
         订单id : Int;
         ab物料 : Int;   // 1A，2B，3不需要
         小钢珠数量 : Int;
         大钢珠数量 : Int;
         存储仓位 : Int;
         当前订单完成 : Bool;
         开始信号 : Int;
         复位信号 : Int;
         订单保留数据 : Array[0..4] of Int;
      END_STRUCT;
   END_VAR
BEGIN
END_DATA_BLOCK

// folder: (top level)

FUNCTION_BLOCK "订单信息下发"   // FB1, LAD
{ S7_Optimized_Access := 'TRUE' }
VERSION : 0.1
   VAR_INPUT
      MES下单请求 : Bool;
      一站可接收 : Int;
      三站已完成 : Int;
   END_VAR
   VAR_OUTPUT
      产线可接收订单 : Bool;
   END_VAR
   VAR
      订单下发步骤 : Int;
      沿 : Bool;
   END_VAR
   VAR_TEMP   // added for the SCL form of the ladder/FBD networks
      _w1 : Bool;
      _w2 : Bool;
   END_VAR
BEGIN

REGION Network 1: 判断三站受否可接单
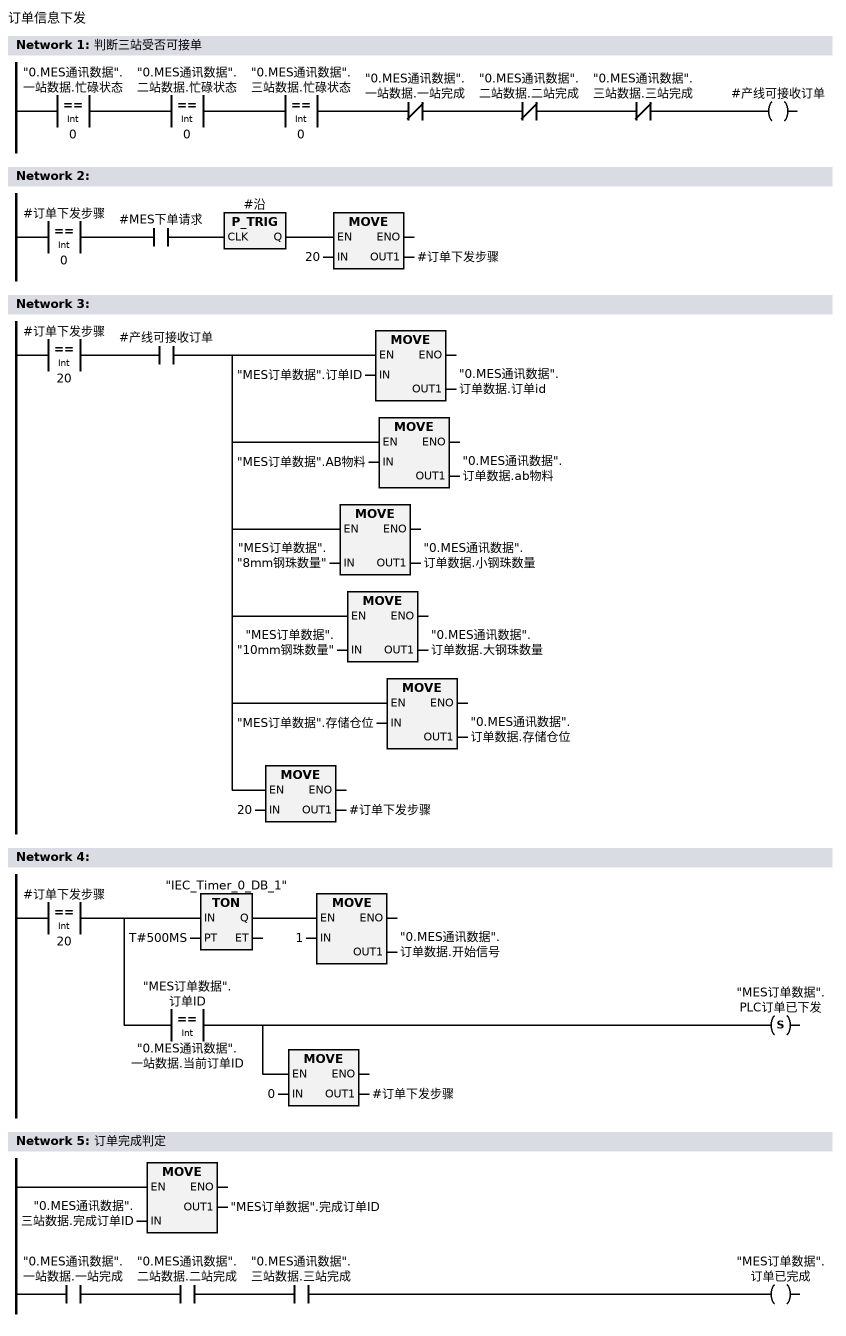
   RUNG wire#powerrail
      { S7_Templates := "SrcType := Int" } EQ_Contact(in1 := "0.MES通讯数据".一站数据.忙碌状态, in2 := 0)
      { S7_Templates := "SrcType := Int" } EQ_Contact(in1 := "0.MES通讯数据".二站数据.忙碌状态, in2 := 0)
      { S7_Templates := "SrcType := Int" } EQ_Contact(in1 := "0.MES通讯数据".三站数据.忙碌状态, in2 := 0)
      I_Contact( "0.MES通讯数据".一站数据.一站完成 )
      I_Contact( "0.MES通讯数据".二站数据.二站完成 )
      I_Contact( "0.MES通讯数据".三站数据.三站完成 )
      Coil( #产线可接收订单 )
   END_RUNG
   // the same network as SCL:
   #产线可接收订单 := ("0.MES通讯数据".一站数据.忙碌状态 = 0) AND ("0.MES通讯数据".二站数据.忙碌状态 = 0) AND ("0.MES通讯数据".三站数据.忙碌状态 = 0) AND NOT "0.MES通讯数据".一站数据.一站完成 AND NOT "0.MES通讯数据".二站数据.二站完成 AND NOT "0.MES通讯数据".三站数据.三站完成;
END_REGION

REGION Network 2
   RUNG wire#powerrail
      { S7_Templates := "SrcType := Int" } EQ_Contact(in1 := #订单下发步骤, in2 := 0)
      Contact( #MES下单请求 )
      P_Trig( #沿 )
      Move(in := 20, out1 => #订单下发步骤)
   END_RUNG
   // the same network as SCL:
   #_w1 := (#订单下发步骤 = 0) AND #MES下单请求;
   #_w2 := #_w1 AND NOT #沿;   // rising edge
   #沿 := #_w1;
   IF #_w2 THEN #订单下发步骤 := 20; END_IF;
END_REGION

REGION Network 3
   RUNG wire#powerrail
      { S7_Templates := "SrcType := Int" } EQ_Contact(in1 := #订单下发步骤, in2 := 20)
      Contact( #产线可接收订单 )
      wire#w1
      Move(in := "MES订单数据".订单ID, out1 => "0.MES通讯数据".订单数据.订单id)
   END_RUNG
   RUNG wire#w1
      Move(in := "MES订单数据".AB物料, out1 => "0.MES通讯数据".订单数据.ab物料)
   END_RUNG
   RUNG wire#w1
      Move(in := "MES订单数据"."8mm钢珠数量", out1 => "0.MES通讯数据".订单数据.小钢珠数量)
   END_RUNG
   RUNG wire#w1
      Move(in := "MES订单数据"."10mm钢珠数量", out1 => "0.MES通讯数据".订单数据.大钢珠数量)
   END_RUNG
   RUNG wire#w1
      Move(in := "MES订单数据".存储仓位, out1 => "0.MES通讯数据".订单数据.存储仓位)
   END_RUNG
   RUNG wire#w1
      Move(in := 20, out1 => #订单下发步骤)
   END_RUNG
   // the same network as SCL:
   IF (#订单下发步骤 = 20) AND #产线可接收订单 THEN
       "0.MES通讯数据".订单数据.订单id := "MES订单数据".订单ID;
       "0.MES通讯数据".订单数据.ab物料 := "MES订单数据".AB物料;
       "0.MES通讯数据".订单数据.小钢珠数量 := "MES订单数据"."8mm钢珠数量";
       "0.MES通讯数据".订单数据.大钢珠数量 := "MES订单数据"."10mm钢珠数量";
       "0.MES通讯数据".订单数据.存储仓位 := "MES订单数据".存储仓位;
       #订单下发步骤 := 20;
   END_IF;
END_REGION

REGION Network 4
   #_w1 := #订单下发步骤 = 20;
   "IEC_Timer_0_DB_1".TON(IN := #_w1, PT := T#500MS);
   IF "IEC_Timer_0_DB_1".Q THEN "0.MES通讯数据".订单数据.开始信号 := 1; END_IF;
   IF #_w1 AND ("MES订单数据".订单ID = "0.MES通讯数据".一站数据.当前订单ID) THEN
       "MES订单数据".PLC订单已下发 := TRUE;
       #订单下发步骤 := 0;
   END_IF;
END_REGION

REGION Network 5: 订单完成判定
   RUNG wire#powerrail
      Move(in := "0.MES通讯数据".三站数据.完成订单ID, out1 => "MES订单数据".完成订单ID)
   END_RUNG
   RUNG wire#powerrail
      Contact( "0.MES通讯数据".一站数据.一站完成 )
      Contact( "0.MES通讯数据".二站数据.二站完成 )
      Contact( "0.MES通讯数据".三站数据.三站完成 )
      Coil( "MES订单数据".订单已完成 )
   END_RUNG
   // the same network as SCL:
   "MES订单数据".完成订单ID := "0.MES通讯数据".三站数据.完成订单ID;
   "MES订单数据".订单已完成 := "0.MES通讯数据".一站数据.一站完成 AND "0.MES通讯数据".二站数据.二站完成 AND "0.MES通讯数据".三站数据.三站完成;
END_REGION
END_FUNCTION_BLOCK

FUNCTION "状态控制" : Void   // FC1, LAD
{ S7_Optimized_Access := 'TRUE' }
VERSION : 0.1
BEGIN

REGION Network 1
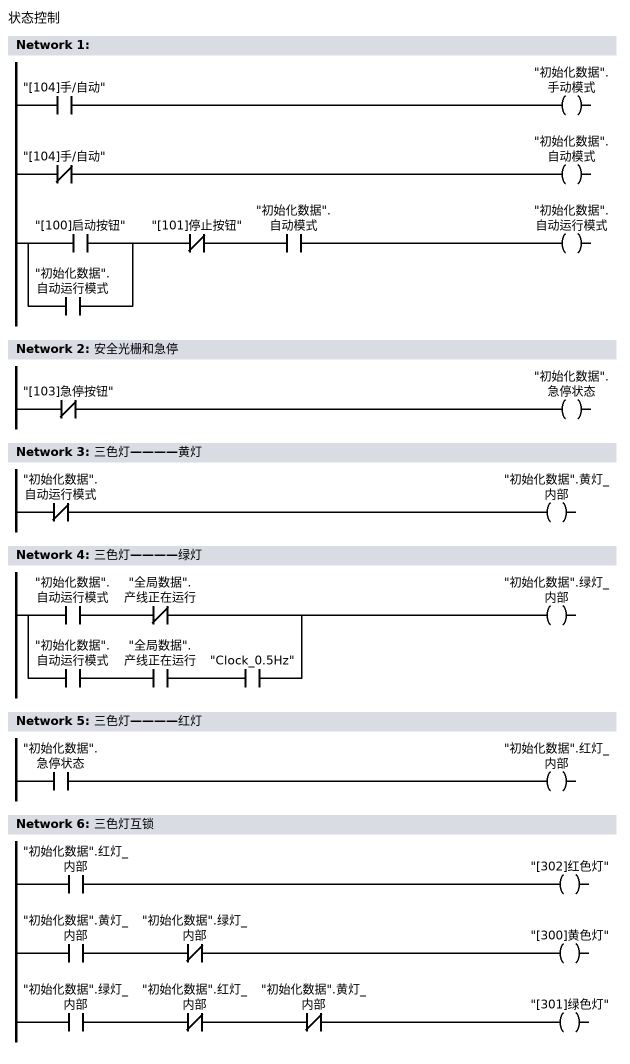
   RUNG wire#powerrail
      Contact( "[104]手/自动" )
      Coil( "初始化数据".手动模式 )
   END_RUNG
   RUNG wire#powerrail
      I_Contact( "[104]手/自动" )
      Coil( "初始化数据".自动模式 )
   END_RUNG
   RUNG wire#powerrail
      Contact( "[100]启动按钮" )
      wire#w1
      I_Contact( "[101]停止按钮" )
      Contact( "初始化数据".自动模式 )
      Coil( "初始化数据".自动运行模式 )
   END_RUNG
   RUNG wire#powerrail
      Contact( "初始化数据".自动运行模式 )
   END_RUNG wire#w1
   // the same network as SCL:
   "初始化数据".手动模式 := "[104]手/自动";
   "初始化数据".自动模式 := NOT "[104]手/自动";
   "初始化数据".自动运行模式 := ("[100]启动按钮" OR "初始化数据".自动运行模式) AND NOT "[101]停止按钮" AND "初始化数据".自动模式;
END_REGION

REGION Network 2: 安全光栅和急停
   RUNG wire#powerrail
      I_Contact( "[103]急停按钮" )
      Coil( "初始化数据".急停状态 )
   END_RUNG
   // the same network as SCL:
   "初始化数据".急停状态 := NOT "[103]急停按钮";
END_REGION

REGION Network 3: 三色灯————黄灯
   RUNG wire#powerrail
      I_Contact( "初始化数据".自动运行模式 )
      Coil( "初始化数据".黄灯_内部 )
   END_RUNG
   // the same network as SCL:
   "初始化数据".黄灯_内部 := NOT "初始化数据".自动运行模式;
END_REGION

REGION Network 4: 三色灯————绿灯
   RUNG wire#powerrail
      Contact( "初始化数据".自动运行模式 )
      I_Contact( "全局数据".产线正在运行 )
      wire#w1
      Coil( "初始化数据".绿灯_内部 )
   END_RUNG
   RUNG wire#powerrail
      Contact( "初始化数据".自动运行模式 )
      Contact( "全局数据".产线正在运行 )
      Contact( "Clock_0.5Hz" )
   END_RUNG wire#w1
   // the same network as SCL:
   "初始化数据".绿灯_内部 := ("初始化数据".自动运行模式 AND NOT "全局数据".产线正在运行) OR ("初始化数据".自动运行模式 AND "全局数据".产线正在运行 AND "Clock_0.5Hz");
END_REGION

REGION Network 5: 三色灯————红灯
   RUNG wire#powerrail
      Contact( "初始化数据".急停状态 )
      Coil( "初始化数据".红灯_内部 )
   END_RUNG
   // the same network as SCL:
   "初始化数据".红灯_内部 := "初始化数据".急停状态;
END_REGION

REGION Network 6: 三色灯互锁
   RUNG wire#powerrail
      Contact( "初始化数据".红灯_内部 )
      Coil( "[302]红色灯" )
   END_RUNG
   RUNG wire#powerrail
      Contact( "初始化数据".黄灯_内部 )
      I_Contact( "初始化数据".绿灯_内部 )
      Coil( "[300]黄色灯" )
   END_RUNG
   RUNG wire#powerrail
      Contact( "初始化数据".绿灯_内部 )
      I_Contact( "初始化数据".红灯_内部 )
      I_Contact( "初始化数据".黄灯_内部 )
      Coil( "[301]绿色灯" )
   END_RUNG
   // the same network as SCL:
   "[302]红色灯" := "初始化数据".红灯_内部;
   "[300]黄色灯" := "初始化数据".黄灯_内部 AND NOT "初始化数据".绿灯_内部;
   "[301]绿色灯" := "初始化数据".绿灯_内部 AND NOT "初始化数据".红灯_内部 AND NOT "初始化数据".黄灯_内部;
END_REGION
END_FUNCTION

FUNCTION "产线复位" : Void   // FC3, LAD
{ S7_Optimized_Access := 'TRUE' }
VERSION : 0.1
BEGIN

REGION Network 1: 产线手动复位
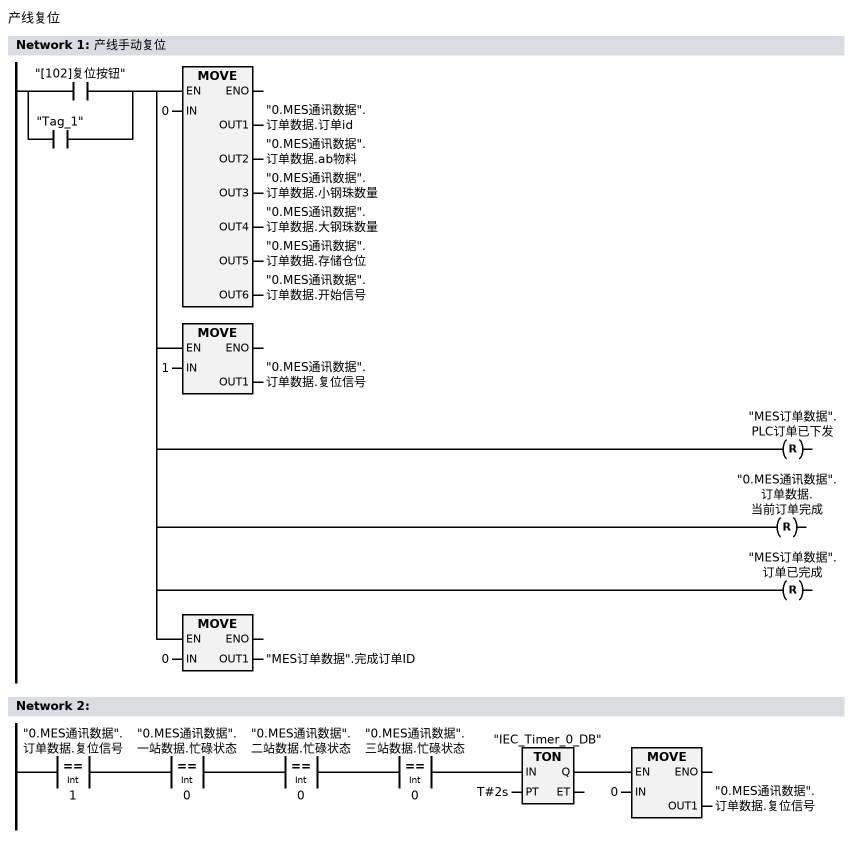
   RUNG wire#powerrail
      Contact( "[102]复位按钮" )
      wire#w1
      Move(in := 0, out1 => "0.MES通讯数据".订单数据.订单id, out2 => "0.MES通讯数据".订单数据.ab物料, out3 => "0.MES通讯数据".订单数据.小钢珠数量, out4 => "0.MES通讯数据".订单数据.大钢珠数量, out5 => "0.MES通讯数据".订单数据.存储仓位, out6 => "0.MES通讯数据".订单数据.开始信号)
   END_RUNG
   RUNG wire#powerrail
      Contact( "Tag_1" )
   END_RUNG wire#w1
   RUNG wire#w1
      Move(in := 1, out1 => "0.MES通讯数据".订单数据.复位信号)
   END_RUNG
   RUNG wire#w1
      R_Coil( "MES订单数据".PLC订单已下发 )
   END_RUNG
   RUNG wire#w1
      R_Coil( "0.MES通讯数据".订单数据.当前订单完成 )
   END_RUNG
   RUNG wire#w1
      R_Coil( "MES订单数据".订单已完成 )
   END_RUNG
   RUNG wire#w1
      Move(in := 0, out1 => "MES订单数据".完成订单ID)
   END_RUNG
   // the same network as SCL:
   IF "[102]复位按钮" OR "Tag_1" THEN
       "0.MES通讯数据".订单数据.订单id := 0;
       "0.MES通讯数据".订单数据.ab物料 := 0;
       "0.MES通讯数据".订单数据.小钢珠数量 := 0;
       "0.MES通讯数据".订单数据.大钢珠数量 := 0;
       "0.MES通讯数据".订单数据.存储仓位 := 0;
       "0.MES通讯数据".订单数据.开始信号 := 0;
       "0.MES通讯数据".订单数据.复位信号 := 1;
       "MES订单数据".PLC订单已下发 := FALSE;
       "0.MES通讯数据".订单数据.当前订单完成 := FALSE;
       "MES订单数据".订单已完成 := FALSE;
       "MES订单数据".完成订单ID := 0;
   END_IF;
END_REGION

REGION Network 2
   "IEC_Timer_0_DB".TON(IN := ("0.MES通讯数据".订单数据.复位信号 = 1) AND ("0.MES通讯数据".一站数据.忙碌状态 = 0) AND ("0.MES通讯数据".二站数据.忙碌状态 = 0) AND ("0.MES通讯数据".三站数据.忙碌状态 = 0),
                        PT := T#2s);
   IF "IEC_Timer_0_DB".Q THEN "0.MES通讯数据".订单数据.复位信号 := 0; END_IF;
END_REGION
END_FUNCTION

FUNCTION "0.MES通讯" : Void   // FC6, LAD
{ S7_Optimized_Access := 'TRUE' }
VERSION : 0.1
BEGIN

REGION Network 1: 心跳
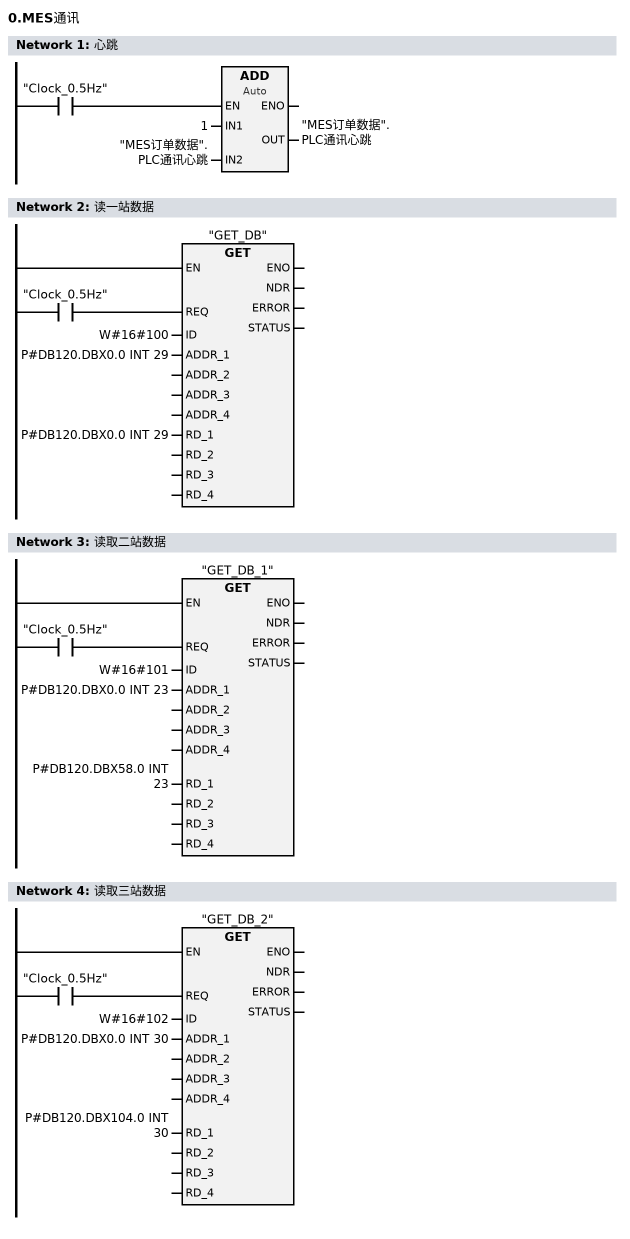
   RUNG wire#powerrail
      Contact( "Clock_0.5Hz" )
      Add(in1 := 1, in2 := "MES订单数据".PLC通讯心跳, out => "MES订单数据".PLC通讯心跳)
   END_RUNG
   // the same network as SCL:
   IF "Clock_0.5Hz" THEN "MES订单数据".PLC通讯心跳 := 1 + "MES订单数据".PLC通讯心跳; END_IF;
END_REGION

REGION Network 2: 读一站数据
   "GET_DB"(REQ := "Clock_0.5Hz",   // GET
            ID := W#16#100,
            ADDR_1 := P#DB120.DBX0.0 INT 29,
            RD_1 := P#DB120.DBX0.0 INT 29);
END_REGION

REGION Network 3: 读取二站数据
   "GET_DB_1"(REQ := "Clock_0.5Hz",   // GET
              ID := W#16#101,
              ADDR_1 := P#DB120.DBX0.0 INT 23,
              RD_1 := P#DB120.DBX58.0 INT 23);
END_REGION

REGION Network 4: 读取三站数据
   "GET_DB_2"(REQ := "Clock_0.5Hz",   // GET
              ID := W#16#102,
              ADDR_1 := P#DB120.DBX0.0 INT 30,
              RD_1 := P#DB120.DBX104.0 INT 30);
END_REGION
END_FUNCTION

ORGANIZATION_BLOCK "Main"   // OB1, LAD, ProgramCycle
TITLE = "Main Program Sweep (Cycle)"
{ S7_Optimized_Access := 'TRUE' }
VERSION : 0.1
   VAR_INPUT
      Initial_Call : Bool;   // Initial call of this OB
      Remanence : Bool;   // =True, if remanent data are available
   END_VAR
   VAR_TEMP   // added for the SCL form of the ladder/FBD networks
      _w1 : Bool;
      _w2 : Bool;
   END_VAR
BEGIN

REGION Network 1: 自动下发订单
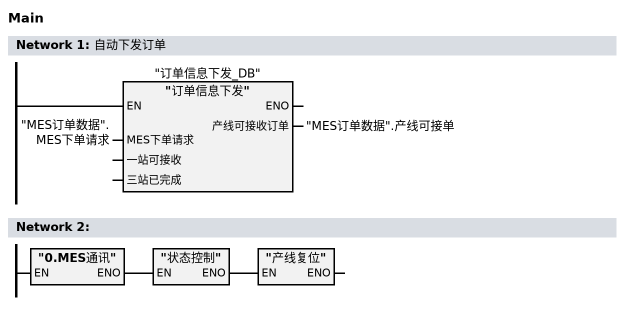
   RUNG wire#powerrail
      "订单信息下发_DB"(MES下单请求 := "MES订单数据".MES下单请求, 一站可接收 :=, 三站已完成 :=, 产线可接收订单 => "MES订单数据".产线可接单)
   END_RUNG
   // the same network as SCL:
   "订单信息下发_DB"(MES下单请求 := "MES订单数据".MES下单请求, 产线可接收订单 => "MES订单数据".产线可接单);   // "订单信息下发"
END_REGION

REGION Network 2
   RUNG wire#powerrail
      "0.MES通讯"()
      "状态控制"()
      "产线复位"()
   END_RUNG
   // the same network as SCL:
   "0.MES通讯"(ENO => #_w1);
   "状态控制"(EN := #_w1, ENO => #_w2);
   IF #_w2 THEN "产线复位"(); END_IF;
END_REGION
END_ORGANIZATION_BLOCK

(* ===== HMI "HMI_RT_1" =====
system functions are stored by id; their names below are inferred from use
connection "HMI_连接_1": ETHERNET, SMART_S7_1200_OMS

HMI tags "默认变量表"
   "[320]底盒推料气缸" : Bool = PLC "[320]底盒推料气缸" AT %Q2.0, 500 ms
   "[112]料仓有无料盒" : Bool = PLC "[112]料仓有无料盒" AT %I1.2, 500 ms
   "[124]推料盒缩回位" : Bool = PLC "[124]推料盒缩回位" AT %I2.4, 500 ms
   "[125]推料盒伸出位" : Bool = PLC "[125]推料盒伸出位" AT %I2.5, 500 ms
   "全局数据块_转盘角度" : Real = PLC 运动控制数据块.转盘目标角度 AT %DB1.DBD0, 1 s
   "全局数据块_转盘设定速度" : Real = PLC 运动控制数据块.转盘目标速度 AT %DB1.DBD4, 1 s
   "[323]取底盒升降气缸" : Bool = PLC "[323]取底盒升降气缸" AT %Q2.3, 1 s
   "[326]取料盒夹爪" : Bool = PLC "[326]取料盒夹爪" AT %Q2.6, 1 s
   "运动控制数据块_机械手实际位置" : Real = PLC 运动控制数据块.机械手实际位置 AT %DB1.DBD26, 1 s
   "运动控制数据块_机械手目标位置" : Real = PLC 运动控制数据块.机械手目标位置 AT %DB1.DBD18, 1 s
   "运动控制数据块_机械手目标速度" : Real = PLC 运动控制数据块.机械手目标速度 AT %DB1.DBD22, 1 s
   "[132]取料盒下降位" : Bool = PLC "[132]取料盒下降位" AT %I3.2, 1 s
   "[133]取料盒上升位" : Bool = PLC "[133]取料盒上升位" AT %I3.3, 1 s
   "[144]机械手夹紧到位" : Bool = PLC "[144]机械手夹紧到位" AT %I4.4, 1 s
   "[145]机械手松开到位" : Bool = PLC "[145]机械手松开到位" AT %I4.5, 1 s
   "[100]伺服左极限" : Bool = PLC "[100]伺服左极限" AT %I0.0, 1 s
   "[101]伺服右极限" : Bool = PLC "[101]伺服右极限" AT %I0.1, 1 s
   "[120]A库物料检测" : Bool = PLC "[120]A库物料检测" AT %I2.0, 1 s
   "[121]B库物料检测" : Bool = PLC "[121]B库物料检测" AT %I2.1, 1 s
   "[126]A推料伸出位" : Bool = PLC "[126]A推料伸出位" AT %I2.6, 1 s
   "[127]A推料缩回位" : Bool = PLC "[127]A推料缩回位" AT %I2.7, 1 s
   "[130]B推料伸出位" : Bool = PLC "[130]B推料伸出位" AT %I3.0, 1 s
   "[131]B推料缩回位" : Bool = PLC "[131]B推料缩回位" AT %I3.1, 1 s
   "[134]取料块伸出位" : Bool = PLC "[134]取料块伸出位" AT %I3.4, 1 s
   "[135]取料块缩回位" : Bool = PLC "[135]取料块缩回位" AT %I3.5, 1 s
   "[136]取料块下降位" : Bool = PLC "[136]取料块下降位" AT %I3.6, 1 s
   "[137]取料块上升位" : Bool = PLC "[137]取料块上升位" AT %I3.7, 1 s
   "[321]A库推料气缸" : Bool = PLC "[321]A库推料气缸" AT %Q2.1, 1 s
   "[322]B库推料气缸" : Bool = PLC "[322]B库推料气缸" AT %Q2.2, 1 s
   "[324]取料块升降气缸" : Bool = PLC "[324]取料块升降气缸" AT %Q2.4, 1 s
   "[325]取料块伸缩气缸" : Bool = PLC "[325]取料块伸缩气缸" AT %Q2.5, 1 s
   "[327]取料块吸盘" : Bool = PLC "[327]取料块吸盘" AT %Q2.7, 1 s
   "[305]转盘皮带电机(正转)" : Bool = PLC "[305]转盘皮带电机(正转)" AT %Q0.5, 1 s
   "[306]转盘皮带电机(反转)" : Bool = PLC "[306]转盘皮带电机(反转)" AT %Q0.6, 1 s
   "运动控制数据块_转盘实际角度" : Real = PLC 运动控制数据块.转盘实际角度 AT %DB1.DBD8, 1 s
   "[310]检测伸缩气缸" : Bool = PLC "[310]检测伸缩气缸" AT %Q1.0, 1 s
   "[311]检测升降气缸" : Bool = PLC "[311]检测升降气缸" AT %Q1.1, 1 s
   "[141]检测缩回位" : Bool = PLC "[141]检测缩回位" AT %I4.1, 1 s
   "[140]检测伸出位" : Bool = PLC "[140]检测伸出位" AT %I4.0, 1 s
   "[142]检测下降位" : Bool = PLC "[142]检测下降位" AT %I4.2, 1 s
   "[143]检测上升位" : Bool = PLC "[143]检测上升位" AT %I4.3, 1 s
   "自动模式数据_当前深度检测" : Real = PLC 自动模式数据.当前深度检测 AT %DB22.DBD42, 1 s
   "运动控制数据块_机械手左移点动" : Bool = PLC 运动控制数据块.机械手左移点动 AT %DB1.DBX35.4, 1 s
   "运动控制数据块_机械手右移点动" : Bool = PLC 运动控制数据块.机械手右移点动 AT %DB1.DBX35.5, 1 s
   "手动模式数据_料块仓选择" : Int = PLC 手动模式数据.料块仓选择 AT %DB12.DBW20, 1 s

screen "推料盒模块" 800x480
   Softkey "Softkey_F1" at 0,0 size 0x0
      on KeyDown: ActivateScreen("推料盒模块", 0)
   Softkey "Softkey_F2" at 0,0 size 0x0
      on KeyDown: ActivateScreen("双供料模块", 0)
   Softkey "Softkey_F3" at 0,0 size 0x0
      on KeyDown: ActivateScreen("双供料模块", 0)
   GraphicView "图形视图_1" at 0,0 size 800x479; Picture "未来智能工厂生产线背景"
   TextField "文本域_6" at 315,21 size 170x37; Text '推料盒模块'
   Button "按钮_2" at 87,403 size 137x60; TextOff '推料盒模块[F1]'
      on Click: ActivateScreen("推料盒模块", 0)
   Button "按钮_3" at 324,403 size 137x60; TextOff '双供料模块[F2]'
      on Click: ActivateScreen("双供料模块", 0)
   Button "按钮_4" at 574,403 size 137x60; TextOff '机械手模块[F3]'
      on Click: ActivateScreen("机械手模块", 0)
   GraphicView "图形视图_2" at 7,88 size 236x306; Picture "图层 1"
   Circle "圆_1" at 702,128 size 31x31
      Appearance <- "[124]推料盒缩回位"
   TextField "文本域_1" at 527,134 size 113x21; Text '推料盒缩回位'
   Circle "圆_2" at 701,165 size 31x31
      Appearance <- "[125]推料盒伸出位"
   TextField "文本域_2" at 526,171 size 113x21; Text '推料盒伸出位'
   Circle "圆_3" at 702,200 size 31x31
      Appearance <- "[112]料仓有无料盒"
   TextField "文本域_4" at 527,209 size 113x21; Text '料仓有无料盒'
   TextField "文本域_5" at 265,134 size 113x21; Text '底盒推料气缸'
   Button "按钮_5" at 382,132 size 57x22; TextOff '置位'
      on Press: SetBit("[320]底盒推料气缸")
   Button "按钮_6" at 446,132 size 57x22; TextOff '复位'
      on Press: ResetBit("[320]底盒推料气缸")
   TextField "文本域_3" at 307,179 size 165x23; Text '旋转皮带步进电机'
   Button "按钮_7" at 261,221 size 81x25; TextOff '正转'
      on Press: SetBit("[305]转盘皮带电机(正转)")
   Button "按钮_8" at 430,221 size 81x25; TextOff '反转'
      on Press: SetBit("[306]转盘皮带电机(反转)")
   IOField "I/O 域_1" at 368,274 size 84x33; FormatPattern 999.99
      ProcessValue <- "运动控制数据块_转盘实际角度"
   TextField "文本域_7" at 313,279 size 65x23; Text '角度：'
   Button "按钮_9" at 346,221 size 81x25; TextOff '停止'
      on Press: ResetBit("[305]转盘皮带电机(正转)"); ResetBit("[306]转盘皮带电机(反转)")
   TextField "文本域_8" at 329,94 size 109x29; Text '输出信号'
   TextField "文本域_9" at 592,94 size 109x29; Text '输入信号'
   TextField "文本域_10" at 261,320 size 113x21; Text '检测伸缩气缸'
   Button "按钮_10" at 378,318 size 57x22; TextOff '置位'
      on Press: SetBit("[310]检测伸缩气缸")
   Button "按钮_11" at 442,318 size 57x22; TextOff '复位'
      on Press: ResetBit("[310]检测伸缩气缸")
   TextField "文本域_11" at 261,352 size 113x21; Text '检测升降气缸'
   Button "按钮_12" at 378,350 size 57x22; TextOff '置位'
      on Press: SetBit("[311]检测升降气缸")
   Button "按钮_13" at 442,350 size 57x22; TextOff '复位'
      on Press: ResetBit("[311]检测升降气缸")
   Circle "圆_4" at 701,237 size 31x31
      Appearance <- "[141]检测缩回位"
   TextField "文本域_12" at 526,245 size 77x21; Text '检测伸出'
   Circle "圆_5" at 653,237 size 31x31
      Appearance <- "[140]检测伸出位"
   TextField "文本域_13" at 526,284 size 77x21; Text '检测下降'
   Circle "圆_6" at 701,276 size 31x31
      Appearance <- "[143]检测上升位"
   Circle "圆_7" at 653,276 size 31x31
      Appearance <- "[142]检测下降位"
   TextField "文本域_14" at 528,327 size 77x21; Text '检测重量'
   IOField "I/O 域_2" at 649,318 size 84x33; FormatPattern 99.99
      ProcessValue <- "自动模式数据_当前深度检测"

screen "双供料模块" 800x480
   Softkey "Softkey_F1" at 0,0 size 0x0
      on KeyDown: ActivateScreen("推料盒模块", 0)
   Softkey "Softkey_F2" at 0,0 size 0x0
      on KeyDown: ActivateScreen("双供料模块", 0)
   Softkey "Softkey_F3" at 0,0 size 0x0
      on KeyDown: ActivateScreen("机械手模块", 0)
   GraphicView "图形视图_1" at 0,0 size 800x479; Picture "未来智能工厂生产线背景"
   Button "按钮_2" at 87,403 size 137x60; TextOff '推料盒模块[F1]'
      on Click: ActivateScreen("推料盒模块", 0)
   Button "按钮_3" at 324,403 size 137x60; TextOff '双供料模块[F2]'
      on Click: ActivateScreen("双供料模块", 0)
   Button "按钮_4" at 574,403 size 137x60; TextOff '机械手模块[F3]'
      on Click: ActivateScreen("机械手模块", 0)
   GraphicView "图形视图_2" at 517,68 size 259x324; Picture "图层 2_1"
   TextField "文本域_3" at 315,14 size 170x37; Text '双供料模块'
   TextField "文本域_11" at 341,77 size 109x29; Text '输入信号'
   TextField "文本域_7" at 287,112 size 123x21; Text 'A料仓有无料块'
   TextField "文本域_12" at 287,145 size 123x21; Text 'B料仓有无料块'
   TextField "文本域_10" at 287,179 size 123x21; Text 'A推料位置检测'
   TextField "文本域_9" at 287,213 size 123x21; Text 'B推料位置检测'
   TextField "文本域_15" at 287,248 size 113x21; Text '取料块伸出位'
   TextField "文本域_16" at 287,282 size 113x21; Text '取料块缩回位'
   TextField "文本域_18" at 287,316 size 113x21; Text '取料块下降位'
   TextField "文本域_17" at 286,350 size 113x21; Text '取料块上升位'
   Circle "圆_9" at 453,345 size 23x23
      Appearance <- "[137]取料块上升位"
   Circle "圆_10" at 453,311 size 23x23
      Appearance <- "[136]取料块下降位"
   Circle "圆_8" at 453,277 size 23x23
      Appearance <- "[135]取料块缩回位"
   Circle "圆_7" at 453,244 size 23x23
      Appearance <- "[134]取料块伸出位"
   Circle "圆_1" at 453,209 size 23x23
      Appearance <- "[131]B推料缩回位"
   Circle "圆_12" at 413,208 size 23x23
      Appearance <- "[130]B推料伸出位"
   Circle "圆_3" at 453,176 size 23x23
      Appearance <- "[127]A推料缩回位"
   Circle "圆_11" at 413,176 size 23x23
      Appearance <- "[126]A推料伸出位"
   Circle "圆_4" at 427,142 size 23x23
      Appearance <- "[121]B库物料检测"
   Circle "圆_2" at 427,108 size 23x23
      Appearance <- "[120]A库物料检测"
   TextField "文本域_8" at 95,71 size 109x29; Text '输出信号'
   TextField "文本域_5" at 19,111 size 105x21; Text 'A库推料气缸'
   Button "按钮_5" at 152,103 size 58x32; TextOff '置位'
      on Press: SetBit("[321]A库推料气缸")
   Button "按钮_6" at 214,103 size 58x32; TextOff '复位'
      on Press: ResetBit("[321]A库推料气缸")
   Button "按钮_8" at 214,159 size 58x32; TextOff '复位'
      on Press: ResetBit("[322]B库推料气缸")
   Button "按钮_7" at 152,159 size 58x32; TextOff '置位'
      on Press: SetBit("[322]B库推料气缸")
   TextField "文本域_1" at 19,167 size 105x21; Text 'B库推料气缸'
   TextField "文本域_2" at 19,224 size 131x21; Text '取料块升降气缸'
   Button "按钮_9" at 152,216 size 58x32; TextOff '置位'
      on Press: SetBit("[324]取料块升降气缸")
   Button "按钮_10" at 214,216 size 58x32; TextOff '复位'
      on Press: ResetBit("[324]取料块升降气缸")
   Button "按钮_12" at 214,272 size 58x32; TextOff '复位'
      on Press: ResetBit("[325]取料块伸缩气缸")
   Button "按钮_11" at 152,272 size 58x32; TextOff '置位'
      on Press: SetBit("[325]取料块伸缩气缸")
   TextField "文本域_4" at 19,280 size 131x21; Text '取料块伸缩气缸'
   TextField "文本域_6" at 19,337 size 95x21; Text '取料块吸盘'
   Button "按钮_13" at 152,329 size 58x32; TextOff '置位'
      on Press: SetBit("[327]取料块吸盘")
   Button "按钮_14" at 214,329 size 58x32; TextOff '复位'
      on Press: ResetBit("[327]取料块吸盘")

screen "机械手模块" 800x480
   Softkey "Softkey_F1" at 0,0 size 0x0
      on KeyDown: ActivateScreen("推料盒模块", 0)
   Softkey "Softkey_F2" at 0,0 size 0x0
      on KeyDown: ActivateScreen("双供料模块", 0)
   Softkey "Softkey_F3" at 0,0 size 0x0
      on KeyDown: ActivateScreen("机械手模块", 0)
   GraphicView "图形视图_1" at 1,0 size 800x479; Picture "未来智能工厂生产线背景"
   Button "按钮_2" at 87,403 size 137x60; TextOff '推料盒模块[F1]'
      on Click: ActivateScreen("推料盒模块", 0)
   Button "按钮_3" at 324,403 size 137x60; TextOff '双供料模块[F2]'
      on Click: ActivateScreen("双供料模块", 0)
   Button "按钮_4" at 574,403 size 137x60; TextOff '机械手模块[F3]'
      on Click: ActivateScreen("机械手模块", 0)
   TextField "文本域_5" at 332,115 size 131x21; Text '取底盒升降气缸'
   Button "按钮_5" at 465,107 size 58x32; TextOff '置位'
      on Press: SetBit("[323]取底盒升降气缸")
   Button "按钮_6" at 527,107 size 58x32; TextOff '复位'
      on Press: ResetBit("[323]取底盒升降气缸")
   TextField "文本域_8" at 403,75 size 109x29; Text '输出信号'
   TextField "文本域_1" at 350,156 size 95x21; Text '取料盒夹爪'
   Button "按钮_7" at 466,148 size 58x32; TextOff '置位'
      on Press: SetBit("[326]取料盒夹爪")
   Button "按钮_8" at 528,148 size 58x32; TextOff '复位'
      on Press: ResetBit("[326]取料盒夹爪")
   TextField "文本域_2" at 413,197 size 77x21; Text '夹爪位置'
   TextField "文本域_7" at 345,230 size 105x23; Text '实际位置：'
   IOField "I/O 域_1" at 458,228 size 97x27; FormatPattern 9999.99
      ProcessValue <- "运动控制数据块_机械手实际位置"
   Button "按钮_9" at 477,345 size 78x32; TextOff '反向移动'
      on Release: ResetBit("运动控制数据块_机械手右移点动")
      on Press: SetBit("运动控制数据块_机械手右移点动")
   Button "按钮_10" at 361,345 size 78x32; TextOff '正向移动'
      on Release: ResetBit("运动控制数据块_机械手左移点动")
      on Press: SetBit("运动控制数据块_机械手左移点动")
   TextField "文本域_4" at 345,265 size 105x23; Text '设定位置：'
   IOField "I/O 域_2" at 458,263 size 97x27; FormatPattern 9999.99
      ProcessValue <- "运动控制数据块_机械手目标位置"
   TextField "文本域_6" at 346,300 size 105x23; Text '设定速度：'
   IOField "I/O 域_3" at 459,298 size 97x27; FormatPattern s999
      ProcessValue <- "运动控制数据块_机械手目标速度"
   TextField "文本域_11" at 654,80 size 109x29; Text '输入信号'
   Circle "圆_2" at 740,110 size 25x25
      Appearance <- "[132]取料盒下降位"
   TextField "文本域_9" at 600,115 size 101x19; Text '取料盒下降位'
   Circle "圆_1" at 740,143 size 25x25
      Appearance <- "[133]取料盒上升位"
   TextField "文本域_10" at 601,148 size 101x19; Text '取料盒上升位'
   Circle "圆_3" at 740,176 size 25x25
      Appearance <- "[144]机械手夹紧到位"
   TextField "文本域_12" at 602,181 size 117x19; Text '机械手夹紧到位'
   Circle "圆_4" at 741,209 size 25x25
      Appearance <- "[145]机械手松开到位"
   TextField "文本域_13" at 602,214 size 117x19; Text '机械手松开到位'
   Circle "圆_5" at 742,242 size 25x25
      Appearance <- "[100]伺服左极限"
   TextField "文本域_14" at 602,247 size 53x19; Text '左极限'
   Circle "圆_6" at 742,274 size 25x25
      Appearance <- "[101]伺服右极限"
   TextField "文本域_15" at 602,279 size 53x19; Text '右极限'
   GraphicView "图形视图_2" at 9,86 size 301x283; Picture "图层 3_1"
   TextField "文本域_3" at 346,18 size 170x37; Text '机械手模块'
   TextField "文本域_16" at 593,325 size 90x20; Text '料块选择：'
   IOField "I/O 域_4" at 683,320 size 99x36; FormatPattern 99
      ProcessValue <- "手动模式数据_料块仓选择"

screen "一站首页" 800x480
   GraphicView "图形视图_1" at 0,0 size 800x479; Picture "未来智能工厂生产线背景"
   Button "按钮_2" at 87,403 size 137x60; TextOff '推料盒模块[F1]'
      on Click: ActivateScreen("推料盒模块", 0)
   Button "按钮_3" at 324,403 size 137x60; TextOff '双供料模块[F2]'
      on Click: ActivateScreen("双供料模块", 0)
   Button "按钮_4" at 574,403 size 137x60; TextOff '机械手模块[F3]'
      on Click: ActivateScreen("机械手模块", 0)
   TextField "文本域_2" at 54,150 size 693x52; Text '非侵入式 AI 智能检测仲裁平台'
   TextField "文本域_1" at 357,244 size 338x40; Text '———自动供料单元'
   Softkey "Softkey_F1" at 0,0 size 0x0
      on KeyDown: ActivateScreen("推料盒模块", 0)
   Softkey "Softkey_F2" at 0,0 size 0x0
      on KeyDown: ActivateScreen("双供料模块", 0)
   Softkey "Softkey_F3" at 0,0 size 0x0
      on KeyDown: ActivateScreen("机械手模块", 0)
*)

(* ===== HMI "HMI_RT_2" =====
system functions are stored by id; their names below are inferred from use
connection "HMI_连接_2": ETHERNET, SMART_S7_1200_OMS

HMI tags "默认变量表"
   "手动模式数据_8mm目标数量" : Int = PLC 手动模式数据.8mm目标数量 AT %DB1.DBW10, 100 ms
   "手动模式数据_10mm目标数量" : Int = PLC 手动模式数据.10mm目标数量 AT %DB1.DBW20, 100 ms
   "手动模式数据_8mm现有钢珠" : Int = PLC 手动模式数据.8mm现有钢珠 AT %DB1.DBW8, 100 ms
   "手动模式数据_10mm现有钢珠" : Int = PLC 手动模式数据.10mm现有钢珠 AT %DB1.DBW18, 100 ms
   "[320]8mm挡停气缸" : Bool = PLC "[320]8mm挡停气缸" AT %Q2.0, 1 s
   "[322]10mm挡停气缸" : Bool = PLC "[322]10mm挡停气缸" AT %Q2.2, 1 s
   "二站数据_电机正转" : Bool = PLC 二站数据.电机正转 AT %DB112.DBX0.4, 1 s
   "[321]8mm推料气缸" : Bool = PLC "[321]8mm推料气缸" AT %Q2.1, 1 s
   "[323]10mm推料气缸" : Bool = PLC "[323]10mm推料气缸" AT %Q2.3, 1 s
   "[124]8mm柱状料仓有无" : Bool = PLC "[124]8mm柱状料仓有无" AT %I2.4, 1 s
   "[131]10mm柱状料仓有无" : Bool = PLC "[131]10mm柱状料仓有无" AT %I3.1, 1 s
   "[105]8mm钢球检测" : Bool = PLC "[105]8mm钢球检测" AT %I0.5, 1 s
   "[106]10mm钢球检测" : Bool = PLC "[106]10mm钢球检测" AT %I0.6, 1 s
   "[120]8mm挡停缩回" : Bool = PLC "[120]8mm挡停缩回" AT %I2.0, 1 s
   "[121]8mm挡停伸出" : Bool = PLC "[121]8mm挡停伸出" AT %I2.1, 1 s
   "[122]8mm料盒到达" : Bool = PLC "[122]8mm料盒到达" AT %I2.2, 1 s
   "[125]10mm挡停缩回" : Bool = PLC "[125]10mm挡停缩回" AT %I2.5, 1 s
   "[126]10mm挡停伸出" : Bool = PLC "[126]10mm挡停伸出" AT %I2.6, 1 s

screen "传送带" 800x480
   GraphicView "图形视图_1" at 0,0 size 800x479; Picture "未来智能工厂生产线背景"
   TextField "文本域_5" at 395,89 size 109x29; Text '输出信号'
   TextField "文本域_6" at 395,139 size 107x21; Text '8mm挡停气缸'
   Button "按钮_8" at 374,169 size 58x32; TextOff '置位'
      on Press: SetBit("[320]8mm挡停气缸")
   Button "按钮_9" at 475,169 size 58x32; TextOff '复位'
      on Press: ResetBit("[320]8mm挡停气缸")
   TextField "文本域_11" at 625,88 size 109x29; Text '输入信号'
   TextField "文本域_7" at 571,133 size 107x21; Text '8mm挡停缩回'
   Circle "圆_2" at 735,126 size 30x30
      Appearance <- "[120]8mm挡停缩回"
   TextField "文本域_9" at 395,204 size 117x21; Text '10mm挡停气缸'
   Button "按钮_10" at 374,234 size 58x32; TextOff '置位'
      on Press: SetBit("[322]10mm挡停气缸")
   Button "按钮_11" at 475,234 size 58x32; TextOff '复位'
      on Press: ResetBit("[322]10mm挡停气缸")
   TextField "文本域_10" at 414,289 size 77x21; Text '皮带控制'
   Button "按钮_12" at 359,319 size 83x32; TextOff '停止'
      on Press: ResetBit("二站数据_电机正转")
   Button "按钮_13" at 460,319 size 83x32; TextOff '启动'
      on Press: SetBit("二站数据_电机正转")
   TextField "文本域_12" at 571,176 size 107x21; Text '8mm挡停伸出'
   Circle "圆_1" at 735,170 size 30x30
      Appearance <- "[121]8mm挡停伸出"
   TextField "文本域_13" at 571,220 size 107x21; Text '8mm料盒到达'
   Circle "圆_3" at 735,214 size 30x30
      Appearance <- "[122]8mm料盒到达"
   TextField "文本域_14" at 571,263 size 117x21; Text '10mm挡停缩回'
   Circle "圆_4" at 735,258 size 30x30
      Appearance <- "[125]10mm挡停缩回"
   TextField "文本域_15" at 571,307 size 117x21; Text '10mm挡停伸出'
   Circle "圆_5" at 735,302 size 30x30
      Appearance <- "[126]10mm挡停伸出"
   TextField "文本域_16" at 571,351 size 117x21; Text '10mm料盒到达'
   Circle "圆_6" at 734,347 size 30x30
      Appearance <- "[122]8mm料盒到达"
   GraphicView "图形视图_3" at 0,105 size 353x267; Picture "图层 6_1"
   TextField "文本域_1" at 315,33 size 170x37; Text '传送带模块'
   Button "按钮_3" at 277,405 size 137x60; TextOff '传送带模块'
      on Click: ActivateScreen("传送带", 0)
   Button "按钮_4" at 461,403 size 137x60; TextOff '灌装模块'
      on Click: ActivateScreen("灌装模块", 0)
   Button "按钮_1" at 94,405 size 137x60; TextOff '首页'
      on Click: ActivateScreen("二站首页", 0)

screen "灌装模块" 800x480
   GraphicView "图形视图_1" at 0,0 size 800x479; Picture "未来智能工厂生产线背景"
   GraphicView "图形视图_4" at 557,88 size 211x317; Picture "图层7_2"
   TextField "文本域_1" at 315,33 size 170x37; Text '供药丸模块'
   TextField "文本域_8" at 126,118 size 109x29; Text '输出信号'
   TextField "文本域_5" at 50,214 size 107x21; Text '8mm推料气缸'
   Button "按钮_8" at 183,206 size 58x32; TextOff '置位'
      on Press: SetBit("[321]8mm推料气缸")
   Button "按钮_9" at 245,206 size 58x32; TextOff '复位'
      on Press: ResetBit("[321]8mm推料气缸")
   Button "按钮_10" at 245,262 size 58x32; TextOff '复位'
      on Press: ResetBit("[323]10mm推料气缸")
   Button "按钮_11" at 183,262 size 58x32; TextOff '置位'
      on Press: SetBit("[323]10mm推料气缸")
   TextField "文本域_2" at 50,270 size 117x21; Text '10mm推料气缸'
   TextField "文本域_11" at 374,124 size 109x29; Text '输入信号'
   TextField "文本域_7" at 330,173 size 143x21; Text '8mm柱状料仓有无'
   TextField "文本域_12" at 330,224 size 153x21; Text '10mm柱状料仓有无'
   TextField "文本域_10" at 330,276 size 107x21; Text '8mm钢球检测'
   TextField "文本域_9" at 330,328 size 117x21; Text '10mm钢球检测'
   Circle "圆_1" at 494,323 size 26x26
      Appearance <- "[106]10mm钢球检测"
   Circle "圆_3" at 496,272 size 26x26
      Appearance <- "[105]8mm钢球检测"
   Circle "圆_4" at 495,222 size 26x26
      Appearance <- "[131]10mm柱状料仓有无"
   Circle "圆_2" at 496,172 size 26x26
      Appearance <- "[124]8mm柱状料仓有无"
   Button "按钮_3" at 277,405 size 137x60; TextOff '传送带模块'
      on Click: ActivateScreen("传送带", 0)
   Button "按钮_4" at 461,403 size 137x60; TextOff '灌装模块'
      on Click: ActivateScreen("灌装模块", 0)
   Button "按钮_1" at 94,405 size 137x60; TextOff '首页'
      on Click: ActivateScreen("二站首页", 0)

screen "二站首页" 800x480
   GraphicView "图形视图_1" at 0,0 size 800x479; Picture "未来智能工厂生产线背景"
   Button "按钮_3" at 163,403 size 137x60; TextOff '传送带模块'
      on Click: ActivateScreen("传送带", 0)
   Button "按钮_4" at 521,403 size 137x60; TextOff '灌装模块'
      on Click: ActivateScreen("灌装模块", 0)
   TextField "文本域_2" at 54,150 size 693x52; Text '非侵入式 AI 智能检测仲裁平台'
   TextField "文本域_1" at 357,244 size 338x40; Text '———智能分拣单元'
*)

(* ===== HMI "HMI_RT_3" =====
system functions are stored by id; their names below are inferred from use
connection "HMI_连接_4": ETHERNET, SMART_S7_1200_OMS

HMI tags "默认变量表"
   "[324]不合格推料气缸" : Bool = PLC "[324]不合格推料气缸" AT %Q2.4, 1 s
   "[320]不合格挡料气缸" : Bool = PLC "[320]不合格挡料气缸" AT %Q2.0, 1 s
   "[311]取料挡料气缸" : Bool = PLC "[311]取料挡料气缸" AT %Q1.1, 1 s
   "全局数据块_变频器启动" : Bool = PLC 全局数据块.变频器启动 AT %DB5.DBX32.0, 1 s
   "[121]不合格挡料伸出位" : Bool = PLC "[121]不合格挡料伸出位" AT %I2.1, 1 s
   "[122]不合格挡料缩回位" : Bool = PLC "[122]不合格挡料缩回位" AT %I2.2, 1 s
   "[120]料盒到位检测" : Bool = PLC "[120]料盒到位检测" AT %I2.0, 1 s
   "[322]滑台移动气缸" : Bool = PLC "[322]滑台移动气缸" AT %Q2.2, 1 s
   "[321滑台伸缩气缸" : Bool = PLC "[321滑台伸缩气缸" AT %Q2.1, 1 s
   "[323]滑台夹爪气缸" : Bool = PLC "[323]滑台夹爪气缸" AT %Q2.3, 1 s
   "[127]滑台夹爪夹紧" : Bool = PLC "[127]滑台夹爪夹紧" AT %I2.7, 1 s
   "[125]]滑台左位" : Bool = PLC "[125]]滑台左位" AT %I2.5, 1 s
   "[126]滑台右位" : Bool = PLC "[126]滑台右位" AT %I2.6, 1 s
   "[130]滑台夹爪松开" : Bool = PLC "[130]滑台夹爪松开" AT %I3.0, 1 s
   "[124]滑台缩回到位" : Bool = PLC "[124]滑台缩回到位" AT %I2.4, 1 s
   "[123]滑台伸出到位" : Bool = PLC "[123]滑台伸出到位" AT %I2.3, 1 s
   "[325]称重抬升气缸" : Bool = PLC "[325]称重抬升气缸" AT %Q2.5, 1 s
   "[326]盒盖推料气缸" : Bool = PLC "[326]盒盖推料气缸" AT %Q2.6, 1 s
   "[330]取盖升降气缸" : Bool = PLC "[330]取盖升降气缸" AT %Q3.0, 1 s
   "[327]取盖伸缩气缸" : Bool = PLC "[327]取盖伸缩气缸" AT %Q2.7, 1 s
   "[331]取盖吸盘" : Bool = PLC "[331]取盖吸盘" AT %Q3.1, 1 s
   "[134]盒盖推料缩回位" : Bool = PLC "[134]盒盖推料缩回位" AT %I3.4, 1 s
   "[133]盒盖推料伸出位" : Bool = PLC "[133]盒盖推料伸出位" AT %I3.3, 1 s
   "[140]取盒盖上升位" : Bool = PLC "[140]取盒盖上升位" AT %I4.0, 1 s
   "[141]取盒盖下降位" : Bool = PLC "[141]取盒盖下降位" AT %I4.1, 1 s
   "[135]取盒盖伸出位" : Bool = PLC "[135]取盒盖伸出位" AT %I3.5, 1 s
   "[136]取盒盖缩回位" : Bool = PLC "[136]取盒盖缩回位" AT %I3.6, 1 s
   "[332]仓储伸缩气缸" : Bool = PLC "[332]仓储伸缩气缸" AT %Q3.2, 1 s
   "[333]仓储升降气缸" : Bool = PLC "[333]仓储升降气缸" AT %Q3.3, 1 s
   "[334]仓储夹爪控制" : Bool = PLC "[334]仓储夹爪控制" AT %Q3.4, 1 s
   "[146]仓储夹爪松开位" : Bool = PLC "[146]仓储夹爪松开位" AT %I4.6, 1 s
   "[145]仓储下降位" : Bool = PLC "[145]仓储下降位" AT %I4.5, 1 s
   "[144]仓储上升位" : Bool = PLC "[144]仓储上升位" AT %I4.4, 1 s
   "[143]仓储缩回位" : Bool = PLC "[143]仓储缩回位" AT %I4.3, 1 s
   "[142]仓储伸出位" : Bool = PLC "[142]仓储伸出位" AT %I4.2, 1 s
   "运动控制数据2_X轴位置" : Real = PLC 运动控制数据2.X轴位置 AT %DB1.DBD0, 1 s
   "运动控制数据2_Y轴位置" : Real = PLC 运动控制数据2.Y轴位置 AT %DB1.DBD4, 1 s

screen "三站首页" 800x480
   GraphicView "图形视图_1" at 0,0 size 800x479; Picture "未来智能工厂生产线背景"
   TextField "文本域_2" at 54,150 size 693x52; Text '非侵入式 AI 智能检测仲裁平台'
   TextField "文本域_1" at 357,244 size 338x40; Text '———智能仓储单元'
   Button "按钮_1" at 18,423 size 133x46; TextOff '首页'
      on Press: ActivateScreen("三站首页", 0)
   Button "按钮_3" at 174,423 size 133x46; TextOff '拍照检测模块'
      on Press: ActivateScreen("0.拍照检测模块", 0)
   Button "按钮_4" at 331,423 size 133x46; TextOff '合格搬运模块'
      on Press: ActivateScreen("1.合格搬运模块", 0)
   Button "按钮_2" at 488,423 size 133x46; TextOff '称重封盖模块'
      on Press: ActivateScreen("2.称重压盖模块", 0)
   Button "按钮_5" at 645,423 size 133x46; TextOff '智能仓储模块'
      on Press: ActivateScreen("3.仓储入库模块", 0)

screen "0.拍照检测模块" 800x480
   GraphicView "图形视图_1" at 0,0 size 800x479; Picture "未来智能工厂生产线背景"
   Button "按钮_1" at 18,423 size 133x46; TextOff '首页'
      on Press: ActivateScreen("三站首页", 0)
   Button "按钮_3" at 174,423 size 133x46; TextOff '拍照检测模块'
      on Press: ActivateScreen("0.拍照检测模块", 0)
   Button "按钮_4" at 331,423 size 133x46; TextOff '合格搬运模块'
      on Press: ActivateScreen("1.合格搬运模块", 0)
   Button "按钮_2" at 488,423 size 133x46; TextOff '称重封盖模块'
      on Press: ActivateScreen("2.称重压盖模块", 0)
   Button "按钮_5" at 645,423 size 133x46; TextOff '智能仓储模块'
      on Press: ActivateScreen("3.仓储入库模块", 0)
   TextField "文本域_1" at 299,17 size 173x31; Text '拍照检测模块'
   GraphicView "图形视图_2" at 570,50 size 211x339; Picture "图层9_1"
   TextField "文本域_8" at 94,69 size 109x29; Text '输出信号'
   TextField "文本域_5" at 21,109 size 131x21; Text '不合格推料气缸'
   Button "按钮_8" at 151,101 size 58x32; TextOff '置位'
      on Press: SetBit("[324]不合格推料气缸")
   Button "按钮_9" at 213,101 size 58x32; TextOff '复位'
      on Press: ResetBit("[324]不合格推料气缸")
   TextField "文本域_11" at 342,67 size 109x29; Text '输入信号'
   TextField "文本域_7" at 288,105 size 95x21; Text '不合格推料'
   Circle "圆_2" at 465,103 size 28x28
      Appearance <- "[122]不合格挡料缩回位"
   TextField "文本域_2" at 22,167 size 131x21; Text '不合格挡料气缸'
   Button "按钮_6" at 152,159 size 58x32; TextOff '置位'
      on Press: SetBit("[320]不合格挡料气缸")
   Button "按钮_7" at 214,159 size 58x32; TextOff '复位'
      on Press: ResetBit("[320]不合格挡料气缸")
   TextField "文本域_3" at 27,225 size 113x21; Text '取料挡料气缸'
   Button "按钮_10" at 152,217 size 58x32; TextOff '置位'
      on Press: SetBit("[311]取料挡料气缸")
   Button "按钮_11" at 214,217 size 58x32; TextOff '复位'
      on Press: ResetBit("[311]取料挡料气缸")
   Circle "圆_1" at 427,103 size 28x28
      Appearance <- "[121]不合格挡料伸出位"
   TextField "文本域_4" at 288,157 size 95x21; Text '不合格挡料'
   Circle "圆_3" at 465,155 size 28x28
      Appearance <- "[122]不合格挡料缩回位"
   Circle "圆_4" at 427,155 size 28x28
      Appearance <- "[121]不合格挡料伸出位"
   TextField "文本域_6" at 288,210 size 113x21; Text '料盒到位检测'
   Circle "圆_5" at 464,208 size 28x28
      Appearance <- "[120]料盒到位检测"
   TextField "文本域_12" at 103,272 size 85x23; Text '皮带控制'
   Button "按钮_12" at 53,303 size 93x37; TextOff '停止'
      on Press: ResetBit("全局数据块_变频器启动")
   Button "按钮_13" at 154,303 size 93x37; TextOff '启动'
      on Press: SetBit("全局数据块_变频器启动")

screen "2.称重压盖模块" 800x480
   GraphicView "图形视图_1" at 0,0 size 800x479; Picture "未来智能工厂生产线背景"
   Button "按钮_1" at 18,423 size 133x46; TextOff '首页'
      on Press: ActivateScreen("三站首页", 0)
   Button "按钮_3" at 174,423 size 133x46; TextOff '拍照检测模块'
      on Press: ActivateScreen("0.拍照检测模块", 0)
   Button "按钮_4" at 331,423 size 133x46; TextOff '合格搬运模块'
      on Press: ActivateScreen("1.合格搬运模块", 0)
   Button "按钮_2" at 488,423 size 133x46; TextOff '称重封盖模块'
      on Press: ActivateScreen("2.称重压盖模块", 0)
   Button "按钮_5" at 645,423 size 133x46; TextOff '智能仓储模块'
      on Press: ActivateScreen("3.仓储入库模块", 0)
   TextField "文本域_1" at 314,20 size 173x31; Text '称重封盖模块'
   GraphicView "图形视图_2" at 20,67 size 213x315; Picture "图层 11"
   TextField "文本域_8" at 370,76 size 109x29; Text '输出信号'
   TextField "文本域_11" at 618,74 size 109x29; Text '输入信号'
   TextField "文本域_7" at 564,115 size 145x23; Text '盒盖推料缩回位'
   Circle "圆_2" at 739,113 size 28x28
      Appearance <- "[134]盒盖推料缩回位"
   TextField "文本域_3" at 294,119 size 113x21; Text '称重抬升气缸'
   Button "按钮_10" at 416,112 size 58x32; TextOff '置位'
      on Press: SetBit("[325]称重抬升气缸")
   Button "按钮_11" at 484,112 size 58x32; TextOff '复位'
      on Press: ResetBit("[325]称重抬升气缸")
   TextField "文本域_2" at 294,171 size 113x21; Text '盒盖推料气缸'
   Button "按钮_6" at 416,164 size 58x32; TextOff '置位'
      on Press: SetBit("[326]盒盖推料气缸")
   Button "按钮_7" at 484,164 size 58x32; TextOff '复位'
      on Press: ResetBit("[326]盒盖推料气缸")
   TextField "文本域_4" at 294,224 size 113x21; Text '取盖升降气缸'
   Button "按钮_8" at 416,217 size 58x32; TextOff '置位'
      on Press: SetBit("[330]取盖升降气缸")
   Button "按钮_9" at 484,217 size 58x32; TextOff '复位'
      on Press: ResetBit("[330]取盖升降气缸")
   TextField "文本域_5" at 294,277 size 113x21; Text '取盖伸缩气缸'
   Button "按钮_12" at 416,269 size 58x32; TextOff '置位'
      on Press: SetBit("[327]取盖伸缩气缸")
   Button "按钮_13" at 484,269 size 58x32; TextOff '复位'
      on Press: ResetBit("[327]取盖伸缩气缸")
   TextField "文本域_6" at 310,330 size 77x21; Text '取盖吸盘'
   Button "按钮_14" at 416,322 size 58x32; TextOff '置位'
      on Press: SetBit("[331]取盖吸盘")
   Button "按钮_15" at 484,322 size 58x32; TextOff '复位'
      on Press: ResetBit("[331]取盖吸盘")
   TextField "文本域_9" at 564,157 size 145x23; Text '盒盖推料伸出位'
   Circle "圆_1" at 739,155 size 28x28
      Appearance <- "[133]盒盖推料伸出位"
   TextField "文本域_10" at 564,199 size 125x23; Text '取盒盖上升位'
   Circle "圆_3" at 739,197 size 28x28
      Appearance <- "[140]取盒盖上升位"
   TextField "文本域_12" at 564,242 size 125x23; Text '取盒盖下降位'
   Circle "圆_4" at 739,240 size 28x28
      Appearance <- "[141]取盒盖下降位"
   TextField "文本域_13" at 564,284 size 125x23; Text '取盒盖伸出位'
   Circle "圆_5" at 739,282 size 28x28
      Appearance <- "[135]取盒盖伸出位"
   TextField "文本域_14" at 564,327 size 125x23; Text '取盒盖缩回位'
   Circle "圆_6" at 739,325 size 28x28
      Appearance <- "[136]取盒盖缩回位"

screen "3.仓储入库模块" 800x480
   GraphicView "图形视图_1" at 0,0 size 800x479; Picture "未来智能工厂生产线背景"
   Button "按钮_1" at 18,423 size 133x46; TextOff '首页'
      on Press: ActivateScreen("三站首页", 0)
   Button "按钮_3" at 174,423 size 133x46; TextOff '拍照检测模块'
      on Press: ActivateScreen("0.拍照检测模块", 0)
   Button "按钮_4" at 331,423 size 133x46; TextOff '合格搬运模块'
      on Press: ActivateScreen("1.合格搬运模块", 0)
   Button "按钮_2" at 488,423 size 133x46; TextOff '称重封盖模块'
      on Press: ActivateScreen("2.称重压盖模块", 0)
   Button "按钮_5" at 645,423 size 133x46; TextOff '智能仓储模块'
      on Press: ActivateScreen("3.仓储入库模块", 0)
   TextField "文本域_1" at 308,19 size 185x33; Text '智能仓储模块'
   GraphicView "图形视图_2" at 488,87 size 307x258; Picture "图层 10"
   TextField "文本域_8" at 91,77 size 109x29; Text '输出信号'
   TextField "文本域_11" at 339,75 size 109x29; Text '输入信号'
   TextField "文本域_7" at 277,105 size 145x23; Text '仓储夹爪松开位'
   Circle "圆_2" at 463,103 size 23x23
      Appearance <- "[146]仓储夹爪松开位"
   TextField "文本域_3" at 15,120 size 113x21; Text '仓储伸缩气缸'
   Button "按钮_10" at 137,113 size 58x32; TextOff '置位'
      on Press: SetBit("[332]仓储伸缩气缸")
   Button "按钮_11" at 205,113 size 58x32; TextOff '复位'
      on Press: ResetBit("[332]仓储伸缩气缸")
   TextField "文本域_2" at 15,156 size 113x21; Text '仓储升降气缸'
   Button "按钮_6" at 137,149 size 58x32; TextOff '置位'
      on Press: SetBit("[333]仓储升降气缸")
   Button "按钮_7" at 205,149 size 58x32; TextOff '复位'
      on Press: ResetBit("[333]仓储升降气缸")
   TextField "文本域_4" at 15,192 size 113x21; Text '仓储夹爪控制'
   Button "按钮_8" at 137,185 size 58x32; TextOff '置位'
      on Press: SetBit("[334]仓储夹爪控制")
   Button "按钮_9" at 205,185 size 58x32; TextOff '复位'
      on Press: ResetBit("[334]仓储夹爪控制")
   TextField "文本域_5" at 97,276 size 69x21; Text 'x轴控制'
   TextField "文本域_6" at 277,128 size 105x23; Text '仓储下降位'
   Circle "圆_1" at 463,126 size 23x23
      Appearance <- "[145]仓储下降位"
   TextField "文本域_9" at 277,151 size 105x23; Text '仓储上升位'
   Circle "圆_3" at 463,149 size 23x23
      Appearance <- "[144]仓储上升位"
   TextField "文本域_10" at 277,173 size 105x23; Text '仓储缩回位'
   Circle "圆_4" at 463,171 size 23x23
      Appearance <- "[143]仓储缩回位"
   TextField "文本域_12" at 277,195 size 105x23; Text '仓储伸出位'
   Circle "圆_5" at 463,193 size 23x23
      Appearance <- "[142]仓储伸出位"
   TextField "文本域_13" at 335,276 size 69x21; Text 'y轴控制'
   TextField "文本域_14" at 24,310 size 105x23; Text '实际位置：'
   IOField "I/O 域_1" at 137,308 size 97x27; FormatPattern s999.99
      ProcessValue <- "运动控制数据2_X轴位置"
   TextField "文本域_15" at 24,345 size 105x23; Text '设定位置：'
   IOField "I/O 域_2" at 137,343 size 97x27; FormatPattern 9999.99
      ProcessValue <- "运动控制数据2_X轴位置"
   TextField "文本域_17" at 292,308 size 105x23; Text '实际位置：'
   IOField "I/O 域_4" at 405,306 size 97x27; FormatPattern s999.99
      ProcessValue <- "运动控制数据2_Y轴位置"
   TextField "文本域_18" at 292,343 size 105x23; Text '设定位置：'
   IOField "I/O 域_5" at 405,341 size 97x27; FormatPattern 9999.99
      ProcessValue <- "运动控制数据2_Y轴位置"

screen "1.合格搬运模块" 800x480
   GraphicView "图形视图_1" at 0,0 size 800x479; Picture "未来智能工厂生产线背景"
   Button "按钮_1" at 18,423 size 133x46; TextOff '首页'
      on Press: ActivateScreen("三站首页", 0)
   Button "按钮_3" at 174,423 size 133x46; TextOff '拍照检测模块'
      on Press: ActivateScreen("0.拍照检测模块", 0)
   Button "按钮_4" at 331,423 size 133x46; TextOff '合格搬运模块'
      on Press: ActivateScreen("1.合格搬运模块", 0)
   Button "按钮_2" at 488,423 size 133x46; TextOff '称重封盖模块'
      on Press: ActivateScreen("2.称重压盖模块", 0)
   Button "按钮_5" at 645,423 size 133x46; TextOff '智能仓储模块'
      on Press: ActivateScreen("3.仓储入库模块", 0)
   TextField "文本域_1" at 314,24 size 173x31; Text '合格搬运模块'
   GraphicView "图形视图_2" at 14,81 size 290x273; Picture "图层8_1"
   TextField "文本域_8" at 384,81 size 109x29; Text '输出信号'
   TextField "文本域_11" at 632,80 size 109x29; Text '输入信号'
   TextField "文本域_7" at 593,139 size 77x21; Text '滑台夹爪'
   Circle "圆_2" at 762,137 size 28x28
      Appearance <- "[130]滑台夹爪松开"
   TextField "文本域_3" at 308,138 size 113x21; Text '取料挡料气缸'
   Button "按钮_10" at 430,131 size 58x32; TextOff '置位'
      on Press: SetBit("[311]取料挡料气缸")
   Button "按钮_11" at 498,131 size 58x32; TextOff '复位'
      on Press: ResetBit("[311]取料挡料气缸")
   Circle "圆_1" at 718,137 size 28x28
      Appearance <- "[127]滑台夹爪夹紧"
   TextField "文本域_2" at 308,179 size 113x21; Text '滑台移动气缸'
   Button "按钮_6" at 430,172 size 58x32; TextOff '置位'
      on Press: SetBit("[322]滑台移动气缸")
   Button "按钮_7" at 498,172 size 58x32; TextOff '复位'
      on Press: ResetBit("[322]滑台移动气缸")
   TextField "文本域_4" at 308,220 size 113x21; Text '滑台伸缩气缸'
   Button "按钮_8" at 430,213 size 58x32; TextOff '置位'
      on Press: SetBit("[321滑台伸缩气缸")
   Button "按钮_9" at 498,213 size 58x32; TextOff '复位'
      on Press: ResetBit("[321滑台伸缩气缸")
   TextField "文本域_5" at 308,261 size 113x21; Text '滑台夹爪气缸'
   Button "按钮_12" at 430,254 size 58x32; TextOff '置位'
      on Press: SetBit("[323]滑台夹爪气缸")
   Button "按钮_13" at 498,254 size 58x32; TextOff '复位'
      on Press: ResetBit("[323]滑台夹爪气缸")
   TextField "文本域_6" at 593,172 size 77x21; Text '滑台位置'
   Circle "圆_3" at 762,170 size 28x28
      Appearance <- "[126]滑台右位"
   Circle "圆_4" at 718,170 size 28x28
      Appearance <- "[125]]滑台左位"
   TextField "文本域_9" at 580,204 size 113x21; Text '滑台缩回到位'
   Circle "圆_5" at 762,204 size 28x28
      Appearance <- "[124]滑台缩回到位"
   TextField "文本域_10" at 580,238 size 113x21; Text '滑台伸出到位'
   Circle "圆_6" at 762,238 size 28x28
      Appearance <- "[123]滑台伸出到位"
*)

(* ===== HMI "HMI_RT_4" =====
system functions are stored by id; their names below are inferred from use
connection "HMI_连接_3": ETHERNET, SMART_S7_1500_OMS

HMI tags "默认变量表"
   "0.MES通讯数据_订单数据_订单id" : Int = PLC "0.MES通讯数据".订单数据.订单id AT %DB120.DBW164, 500 ms
   "0.MES通讯数据_订单数据_ab物料" : Int = PLC "0.MES通讯数据".订单数据.ab物料 AT %DB120.DBW166, 500 ms
   "0.MES通讯数据_订单数据_小钢珠数量" : Int = PLC "0.MES通讯数据".订单数据.小钢珠数量 AT %DB120.DBW168, 500 ms
   "0.MES通讯数据_订单数据_大钢珠数量" : Int = PLC "0.MES通讯数据".订单数据.大钢珠数量 AT %DB120.DBW170, 500 ms
   "0.MES通讯数据_订单数据_存储仓位" : Int = PLC "0.MES通讯数据".订单数据.存储仓位 AT %DB120.DBW172, 500 ms
   "0.MES通讯数据_订单数据_复位信号" : Int = PLC "0.MES通讯数据".订单数据.复位信号 AT %DB120.DBW178, 500 ms
   "0.MES通讯数据_订单数据_开始信号" : Int = PLC "0.MES通讯数据".订单数据.开始信号 AT %DB120.DBW176, 500 ms
   "全局数据_触摸屏下单按钮" : Bool = PLC 全局数据.触摸屏下单按钮 AT %DB3.DBX0.3, 100 ms
   "全局数据_触摸屏复位按钮" : Bool = PLC 全局数据.触摸屏复位按钮 AT %DB3.DBX0.4, 100 ms

screen "下单界面" 800x480
   GraphicView "图形视图_1" at 0,0 size 800x479; Picture "未来智能工厂生产线背景"
   Button "按钮_1" at 580,314 size 119x61; TextOff '下单'
      on Press: SetBit("全局数据_触摸屏下单按钮")
      on Release: ResetBit("全局数据_触摸屏下单按钮")
   TextField "文本域_1" at 487,182 size 125x27; Text '大钢珠数量'
   TextField "文本域_2" at 146,188 size 125x27; Text '小钢珠数量'
   TextField "文本域_3" at 498,86 size 101x27; Text '料块种类'
   TextField "文本域_4" at 158,284 size 101x27; Text '入库仓位'
   IOField "I/O 域_1" at 495,130 size 104x41; FormatPattern 99
      ProcessValue <- "0.MES通讯数据_订单数据_ab物料"
   IOField "I/O 域_2" at 157,227 size 104x41; FormatPattern 99
      ProcessValue <- "0.MES通讯数据_订单数据_小钢珠数量"
   IOField "I/O 域_3" at 498,227 size 104x41; FormatPattern 99
      ProcessValue <- "0.MES通讯数据_订单数据_大钢珠数量"
   IOField "I/O 域_4" at 157,326 size 104x41; FormatPattern 99
      ProcessValue <- "0.MES通讯数据_订单数据_存储仓位"
   TextField "文本域_5" at 169,86 size 79x27; Text '订单ID'
   IOField "I/O 域_5" at 157,130 size 104x41; FormatPattern 999999
      ProcessValue <- "0.MES通讯数据_订单数据_订单id"
   Button "按钮_2" at 404,311 size 115x64; TextOff '设备复位'
      on Press: SetBit("全局数据_触摸屏复位按钮")
      on Release: ResetBit("全局数据_触摸屏复位按钮")
   TextField "文本域_6" at 332,26 size 137x37; Text '下单界面'
   Button "按钮_3" at 174,425 size 133x46; TextOff '首页'
      on Press: ActivateScreen("首页", 0)
   Button "按钮_4" at 330,425 size 133x46; TextOff '手动下单'
      on Press: ActivateScreen("首页", 0)
   Button "按钮_5" at 487,425 size 133x46; TextOff '数据检测'
      on Press: ActivateScreen("首页", 0)

screen "首页" 800x480
   GraphicView "图形视图_1" at 0,0 size 800x479; Picture "未来智能工厂生产线背景"
   TextField "文本域_2" at 54,150 size 693x52; Text '非侵入式 AI 智能检测仲裁平台'
   TextField "文本域_1" at 357,244 size 338x40; Text '———数据管理单元'
   Button "按钮_1" at 174,425 size 133x46; TextOff '首页'
      on Press: ActivateScreen("首页", 0)
   Button "按钮_3" at 330,425 size 133x46; TextOff '手动下单'
      on Press: ActivateScreen("首页", 0)
   Button "按钮_4" at 487,425 size 133x46; TextOff '数据检测'
      on Press: ActivateScreen("首页", 0)
*)